  MoveL 521 to (0, -31.79, 55.65) mm, rotated rx 170.45 ry 0 rz 180 deg; joints [-13.216, -55.69, 111.554, 164.16, 56.887, -90.738]
  MoveL 522 to (-200, -31.79, 55.65) mm, rotated rx 170.45 ry 0 rz 180 deg; joints [-15.372, -64.732, 127.633, 162.838, 63.944, -91.824]
  MoveL 523 to (-200, -32.38, 55.53) mm, rotated rx 167.27 ry 0 rz 180 deg; joints [-15.299, -65.985, 127.45, 162.704, 62.564, -94.567]
  MoveL 524 to (0, -32.38, 55.53) mm, rotated rx 167.27 ry 0 rz 180 deg; joints [-13.153, -56.711, 111.391, 164.018, 55.738, -93.573]
  MoveL 525 to (0, -32.96, 55.39) mm, rotated rx 164.09 ry 0 rz 180 deg; joints [-13.044, -57.718, 111.217, 163.922, 54.585, -96.433]
  MoveL 526 to (-200, -32.96, 55.39) mm, rotated rx 164.09 ry 0 rz 180 deg; joints [-15.175, -67.219, 127.255, 162.616, 61.181, -97.333]
  MoveL 527 to (-200, -33.53, 55.21) mm, rotated rx 160.9 ry 0 rz 180 deg; joints [-14.999, -68.432, 127.047, 162.576, 59.799, -100.128]
  MoveL 528 to (0, -33.53, 55.21) mm, rotated rx 160.9 ry 0 rz 180 deg; joints [-12.891, -58.708, 111.032, 163.872, 53.431, -99.324]
  MoveL 529 to (0, -34.09, 54.99) mm, rotated rx 157.72 ry 0 rz 180 deg; joints [-12.693, -59.678, 110.838, 163.872, 52.279, -102.249]
  MoveL 530 to (-200, -34.09, 54.99) mm, rotated rx 157.72 ry 0 rz 180 deg; joints [-14.771, -69.618, 126.828, 162.586, 58.422, -102.955]
  MoveL 531 to (-200, -34.64, 54.75) mm, rotated rx 154.53 ry 0 rz 180 deg; joints [-14.492, -70.775, 126.599, 162.65, 57.053, -105.822]
  MoveL 532 to (0, -34.64, 54.75) mm, rotated rx 154.53 ry 0 rz 180 deg; joints [-12.451, -60.626, 110.636, 163.924, 51.131, -105.214]
  MoveL 533 to (0, -35.18, 54.48) mm, rotated rx 151.35 ry 0 rz 180 deg; joints [-12.165, -61.547, 110.426, 164.031, 49.993, -108.224]
  MoveL 534 to (-200, -35.18, 54.48) mm, rotated rx 151.35 ry 0 rz 180 deg; joints [-14.163, -71.9, 126.361, 162.77, 55.696, -108.734]
  MoveL 535 to (-200, -35.7, 54.18) mm, rotated rx 148.17 ry 0 rz 180 deg; joints [-13.784, -72.989, 126.115, 162.95, 54.354, -111.698]
  MoveL 536 to (0, -35.7, 54.18) mm, rotated rx 148.17 ry 0 rz 180 deg; joints [-11.836, -62.442, 110.21, 164.197, 48.865, -111.284]
  MoveL 537 to (0, -36.2, 53.84) mm, rotated rx 144.99 ry 0 rz 180 deg; joints [-11.464, -63.305, 109.989, 164.425, 47.752, -114.399]
  MoveL 538 to (-200, -36.2, 53.84) mm, rotated rx 144.99 ry 0 rz 180 deg; joints [-13.356, -74.041, 125.863, 163.195, 53.031, -114.72]
  MoveL 539 to (-200, -36.68, 53.49) mm, rotated rx 141.8 ry 0 rz 180 deg; joints [-12.879, -75.052, 125.607, 163.507, 51.731, -117.806]
  MoveL 540 to (0, -36.68, 53.49) mm, rotated rx 141.8 ry 0 rz 180 deg; joints [-11.052, -64.137, 109.764, 164.717, 46.658, -117.575]
  MoveL 541 to (0, -37.14, 53.1) mm, rotated rx 138.62 ry 0 rz 180 deg; joints [-10.598, -64.933, 109.536, 165.079, 45.585, -120.816]
  MoveL 542 to (-200, -37.14, 53.1) mm, rotated rx 138.62 ry 0 rz 180 deg; joints [-12.355, -76.019, 125.348, 163.891, 50.459, -120.962]
  MoveL 543 to (-200, -37.58, 52.7) mm, rotated rx 135.44 ry 0 rz 180 deg; joints [-11.785, -76.941, 125.087, 164.352, 49.218, -124.195]
  MoveL 544 to (0, -37.58, 52.7) mm, rotated rx 135.44 ry 0 rz 180 deg; joints [-10.105, -65.693, 109.307, 165.513, 44.539, -124.128]
  MoveL 545 to (0, -37.99, 52.26) mm, rotated rx 132.25 ry 0 rz 180 deg; joints [-9.574, -66.415, 109.079, 166.023, 43.523, -127.516]
  MoveL 546 to (-200, -37.99, 52.26) mm, rotated rx 132.25 ry 0 rz 180 deg; joints [-11.17, -77.816, 124.826, 164.893, 48.014, -127.51]
  MoveL 547 to (-200, -38.38, 51.81) mm, rotated rx 129.07 ry 0 rz 180 deg; joints [-10.512, -78.64, 124.568, 165.519, 46.851, -130.914]
  MoveL 548 to (0, -38.38, 51.81) mm, rotated rx 129.07 ry 0 rz 180 deg; joints [-9.006, -67.096, 108.852, 166.613, 42.541, -130.984]
  MoveL 549 to (0, -38.75, 51.33) mm, rotated rx 125.89 ry 0 rz 180 deg; joints [-8.403, -67.735, 108.628, 167.284, 41.598, -134.535]
  MoveL 550 to (-200, -38.75, 51.33) mm, rotated rx 125.89 ry 0 rz 180 deg; joints [-9.811, -79.413, 124.313, 166.234, 45.735, -134.409]
  MoveL 551 to (-200, -39.09, 50.84) mm, rotated rx 122.7 ry 0 rz 180 deg; joints [-9.071, -80.133, 124.064, 167.04, 44.67, -138.001]
  MoveL 552 to (0, -39.09, 50.84) mm, rotated rx 122.7 ry 0 rz 180 deg; joints [-7.766, -68.33, 108.408, 168.04, 40.698, -138.172]
  MoveL 553 to (0, -39.4, 50.32) mm, rotated rx 119.52 ry 0 rz 180 deg; joints [-7.098, -68.881, 108.194, 168.881, 39.847, -141.898]
  MoveL 554 to (-200, -39.4, 50.32) mm, rotated rx 119.52 ry 0 rz 180 deg; joints [-8.293, -80.797, 123.822, 167.941, 43.662, -141.693]
  MoveL 555 to (-200, -39.68, 49.79) mm, rotated rx 116.34 ry 0 rz 180 deg; joints [-7.48, -81.406, 123.588, 168.937, 42.718, -145.487]
  MoveL 556 to (0, -39.68, 49.79) mm, rotated rx 116.34 ry 0 rz 180 deg; joints [-6.399, -69.385, 107.988, 169.809, 39.048, -145.714]
  MoveL 557 to (0, -39.93, 49.25) mm, rotated rx 113.16 ry 0 rz 180 deg; joints [-5.673, -69.842, 107.79, 170.823, 38.306, -149.62]
  MoveL 558 to (-200, -39.93, 49.25) mm, rotated rx 113.16 ry 0 rz 180 deg; joints [-6.633, -81.956, 123.364, 170.028, 41.841, -149.382]
  MoveL 559 to (-200, -40.15, 48.69) mm, rotated rx 109.97 ry 0 rz 180 deg; joints [-5.756, -82.448, 123.153, 171.213, 41.039, -153.378]
  MoveL 560 to (0, -40.15, 48.69) mm, rotated rx 109.97 ry 0 rz 180 deg; joints [-4.922, -70.251, 107.602, 171.922, 37.627, -153.614]
  MoveL 561 to (0, -40.34, 48.12) mm, rotated rx 106.79 ry 0 rz 180 deg; joints [-4.147, -70.61, 107.424, 173.101, 37.014, -157.692]
  MoveL 562 to (-200, -40.34, 48.12) mm, rotated rx 106.79 ry 0 rz 180 deg; joints [-4.852, -82.881, 122.954, 172.489, 40.317, -157.47]
  MoveL 563 to (-200, -40.5, 47.54) mm, rotated rx 103.61 ry 0 rz 180 deg; joints [-3.922, -83.252, 122.77, 173.85, 39.68, -161.653]
  MoveL 564 to (0, -40.5, 47.54) mm, rotated rx 103.61 ry 0 rz 180 deg; joints [-3.352, -70.919, 107.259, 174.355, 36.473, -161.85]
  MoveL 565 to (0, -40.62, 46.95) mm, rotated rx 100.42 ry 0 rz 180 deg; joints [-2.539, -71.178, 107.107, 175.679, 36.006, -166.079]
  MoveL 566 to (-200, -40.62, 46.95) mm, rotated rx 100.42 ry 0 rz 180 deg; joints [-2.971, -83.563, 122.601, 175.289, 39.133, -165.919]
  MoveL 567 to (-200, -40.71, 46.36) mm, rotated rx 97.24 ry 0 rz 180 deg; joints [-2.002, -83.812, 122.449, 176.795, 38.681, -170.258]
  MoveL 568 to (0, -40.71, 46.36) mm, rotated rx 97.24 ry 0 rz 180 deg; joints [-1.711, -71.386, 106.969, 177.062, 35.619, -170.372]
  MoveL 569 to (0, -40.77, 45.76) mm, rotated rx 94.06 ry 0 rz 180 deg; joints [-0.87, -71.542, 106.846, 178.494, 35.313, -174.715]
  MoveL 570 to (-200, -40.77, 45.76) mm, rotated rx 94.06 ry 0 rz 180 deg; joints [-1.019, -83.999, 122.314, 178.357, 38.327, -174.655]
  MoveL 571 to (-200, -40.8, 45.16) mm, rotated rx 90.87 ry 0 rz 180 deg; joints [-0.024, -84.123, 122.198, 179.961, 38.074, -179.096]
  MoveL 572 to (0, -40.8, 45.16) mm, rotated rx 90.87 ry 0 rz 180 deg; joints [-0.021, -71.646, 106.738, 179.964, 35.092, -179.097]
  MoveL 573 to (0, -40.8, 44.56) mm, rotated rx 90 ry 0 rz 180 deg; joints [0.232, -71.666, 106.711, -179.597, 35.046, 179.67]
  MoveL 574 to (-200, -40.8, 44.56) mm, rotated rx 90 ry 0 rz 180 deg; joints [0.271, -84.147, 122.169, -179.56, 38.023, 179.653]
  MoveL 575 to (-200, -40.8, 43.97) mm, rotated rx 90 ry 0 rz 180 deg; joints [0.301, -84.146, 122.169, -179.512, 38.023, 179.616]
  MoveL 576 to (0, -40.8, 43.97) mm, rotated rx 90 ry 0 rz 180 deg; joints [0.257, -71.666, 106.711, -179.553, 35.046, 179.634]
  MoveL 577 to (0, -40.8, 43.37) mm, rotated rx 90 ry 0 rz 180 deg; joints [0.282, -71.665, 106.711, -179.509, 35.046, 179.598]
  MoveL 578 to (-200, -40.8, 43.37) mm, rotated rx 90 ry 0 rz 180 deg; joints [0.33, -84.146, 122.169, -179.464, 38.024, 179.578]
  MoveL 579 to (-200, -40.8, 42.77) mm, rotated rx 90 ry 0 rz 180 deg; joints [0.359, -84.146, 122.168, -179.417, 38.024, 179.541]
  MoveL 580 to (0, -40.8, 42.77) mm, rotated rx 90 ry 0 rz 180 deg; joints [0.307, -71.665, 106.71, -179.466, 35.046, 179.562]
  MoveL 581 to (0, -40.8, 42.16) mm, rotated rx 90 ry 0 rz 180 deg; joints [0.332, -71.665, 106.71, -179.422, 35.046, 179.527]
  MoveL 582 to (-200, -40.8, 42.16) mm, rotated rx 90 ry 0 rz 180 deg; joints [0.389, -84.146, 122.168, -179.369, 38.024, 179.503]
  MoveL 583 to (-200, -40.8, 41.56) mm, rotated rx 90 ry 0 rz 180 deg; joints [0.418, -84.145, 122.168, -179.322, 38.024, 179.466]
  MoveL 584 to (0, -40.8, 41.56) mm, rotated rx 90 ry 0 rz 180 deg; joints [0.357, -71.665, 106.71, -179.378, 35.047, 179.491]
  MoveL 585 to (0, -40.8, 40.97) mm, rotated rx 90 ry 0 rz 180 deg; joints [0.382, -71.665, 106.709, -179.335, 35.047, 179.455]
  MoveL 586 to (-200, -40.8, 40.97) mm, rotated rx 90 ry 0 rz 180 deg; joints [0.447, -84.145, 122.167, -179.274, 38.025, 179.428]
  MoveL 587 to (-200, -40.8, 40.37) mm, rotated rx 90 ry 0 rz 180 deg; joints [0.477, -84.145, 122.167, -179.226, 38.025, 179.391]
  MoveL 588 to (0, -40.8, 40.37) mm, rotated rx 90 ry 0 rz 180 deg; joints [0.407, -71.664, 106.709, -179.291, 35.047, 179.42]
  MoveL 589 to (0, -40.8, 39.77) mm, rotated rx 90 ry 0 rz 180 deg; joints [0.432, -71.664, 106.709, -179.247, 35.047, 179.384]
  MoveL 590 to (-200, -40.8, 39.77) mm, rotated rx 90 ry 0 rz 180 deg; joints [0.506, -84.144, 122.167, -179.179, 38.025, 179.353]
  MoveL 591 to (-200, -40.8, 39.16) mm, rotated rx 90 ry 0 rz 180 deg; joints [0.535, -84.144, 122.166, -179.131, 38.025, 179.316]
  MoveL 592 to (0, -40.8, 39.16) mm, rotated rx 90 ry 0 rz 180 deg; joints [0.457, -71.664, 106.708, -179.204, 35.047, 179.348]
  MoveL 593 to (0, -40.8, 38.56) mm, rotated rx 90 ry 0 rz 180 deg; joints [0.482, -71.663, 106.708, -179.16, 35.047, 179.312]
  MoveL 594 to (-200, -40.8, 38.56) mm, rotated rx 90 ry 0 rz 180 deg; joints [0.565, -84.144, 122.166, -179.084, 38.026, 179.278]
  MoveL 595 to (-200, -40.8, 37.97) mm, rotated rx 90 ry 0 rz 180 deg; joints [0.594, -84.143, 122.165, -179.036, 38.026, 179.241]
  MoveL 596 to (0, -40.8, 37.97) mm, rotated rx 90 ry 0 rz 180 deg; joints [0.507, -71.663, 106.708, -179.117, 35.048, 179.277]
  MoveL 597 to (0, -40.8, 37.37) mm, rotated rx 90 ry 0 rz 180 deg; joints [0.532, -71.663, 106.707, -179.073, 35.048, 179.241]
  MoveL 598 to (-200, -40.8, 37.37) mm, rotated rx 90 ry 0 rz 180 deg; joints [0.623, -84.143, 122.165, -178.988, 38.026, 179.203]
  MoveL 599 to (-200, -40.8, 36.77) mm, rotated rx 90 ry 0 rz 180 deg; joints [0.653, -84.143, 122.165, -178.941, 38.027, 179.166]
  MoveL 600 to (0, -40.8, 36.77) mm, rotated rx 90 ry 0 rz 180 deg; joints [0.557, -71.662, 106.707, -179.029, 35.048, 179.205]
  MoveL 601 to (0, -40.8, 36.16) mm, rotated rx 90 ry 0 rz 180 deg; joints [0.582, -71.662, 106.706, -178.986, 35.048, 179.17]
  MoveL 602 to (-200, -40.8, 36.16) mm, rotated rx 90 ry 0 rz 180 deg; joints [0.682, -84.142, 122.164, -178.893, 38.027, 179.128]
  MoveL 603 to (-200, -40.8, 35.56) mm, rotated rx 90 ry 0 rz 180 deg; joints [0.711, -84.142, 122.163, -178.845, 38.028, 179.091]
  MoveL 604 to (0, -40.8, 35.56) mm, rotated rx 90 ry 0 rz 180 deg; joints [0.608, -71.662, 106.706, -178.942, 35.048, 179.134]
  MoveL 605 to (0, -40.8, 34.97) mm, rotated rx 90 ry 0 rz 180 deg; joints [0.633, -71.661, 106.705, -178.898, 35.049, 179.098]
  MoveL 606 to (-200, -40.8, 34.97) mm, rotated rx 90 ry 0 rz 180 deg; joints [0.741, -84.141, 122.163, -178.798, 38.028, 179.053]
  MoveL 607 to (-200, -40.8, 34.37) mm, rotated rx 90 ry 0 rz 180 deg; joints [0.77, -84.141, 122.162, -178.75, 38.028, 179.016]
  MoveL 608 to (0, -40.8, 34.37) mm, rotated rx 90 ry 0 rz 180 deg; joints [0.658, -71.661, 106.704, -178.855, 35.049, 179.062]
  MoveL 609 to (0, -40.8, 33.77) mm, rotated rx 90 ry 0 rz 180 deg; joints [0.683, -71.66, 106.704, -178.811, 35.049, 179.027]
  MoveL 610 to (-200, -40.8, 33.77) mm, rotated rx 90 ry 0 rz 180 deg; joints [0.799, -84.14, 122.162, -178.703, 38.029, 178.978]
  MoveL 611 to (-200, -40.8, 33.16) mm, rotated rx 90 ry 0 rz 180 deg; joints [0.829, -84.14, 122.161, -178.655, 38.029, 178.941]
  MoveL 612 to (0, -40.8, 33.16) mm, rotated rx 90 ry 0 rz 180 deg; joints [0.708, -71.66, 106.703, -178.768, 35.05, 178.991]
  MoveL 613 to (0, -40.8, 32.56) mm, rotated rx 90 ry 0 rz 180 deg; joints [0.733, -71.66, 106.703, -178.724, 35.05, 178.955]
  MoveL 614 to (-200, -40.8, 32.56) mm, rotated rx 90 ry 0 rz 180 deg; joints [0.858, -84.139, 122.161, -178.607, 38.03, 178.903]
  MoveL 615 to (-200, -40.8, 31.96) mm, rotated rx 90 ry 0 rz 180 deg; joints [0.887, -84.138, 122.16, -178.56, 38.03, 178.866]
  MoveL 616 to (0, -40.8, 31.96) mm, rotated rx 90 ry 0 rz 180 deg; joints [0.758, -71.659, 106.702, -178.68, 35.05, 178.92]
  MoveL 617 to (0, -40.8, 31.36) mm, rotated rx 90 ry 0 rz 180 deg; joints [0.783, -71.659, 106.701, -178.637, 35.05, 178.884]
  MoveL 618 to (-200, -40.8, 31.36) mm, rotated rx 90 ry 0 rz 180 deg; joints [0.916, -84.138, 122.159, -178.512, 38.031, 178.828]
  MoveL 619 to (-200, -40.8, 30.77) mm, rotated rx 90 ry 0 rz 180 deg; joints [0.946, -84.137, 122.158, -178.465, 38.031, 178.791]
  MoveL 620 to (0, -40.8, 30.77) mm, rotated rx 90 ry 0 rz 180 deg; joints [0.808, -71.658, 106.701, -178.593, 35.051, 178.848]
  MoveL 621 to (0, -40.8, 30.16) mm, rotated rx 90 ry 0 rz 180 deg; joints [0.833, -71.657, 106.7, -178.549, 35.051, 178.812]
  MoveL 622 to (-200, -40.8, 30.16) mm, rotated rx 90 ry 0 rz 180 deg; joints [0.975, -84.136, 122.158, -178.417, 38.032, 178.753]
  MoveL 623 to (-200, -40.8, 29.57) mm, rotated rx 90 ry 0 rz 180 deg; joints [1.004, -84.136, 122.157, -178.37, 38.032, 178.716]
  MoveL 624 to (0, -40.8, 29.57) mm, rotated rx 90 ry 0 rz 180 deg; joints [0.858, -71.657, 106.699, -178.506, 35.051, 178.777]
  MoveL 625 to (0, -40.8, 28.96) mm, rotated rx 90 ry 0 rz 180 deg; joints [0.883, -71.656, 106.698, -178.462, 35.052, 178.741]
  MoveL 626 to (-200, -40.8, 28.96) mm, rotated rx 90 ry 0 rz 180 deg; joints [1.034, -84.135, 122.156, -178.322, 38.033, 178.678]
  MoveL 627 to (-200, -40.8, 28.36) mm, rotated rx 90 ry 0 rz 180 deg; joints [1.063, -84.134, 122.155, -178.274, 38.034, 178.641]
  MoveL 628 to (0, -40.8, 28.36) mm, rotated rx 90 ry 0 rz 180 deg; joints [0.908, -71.656, 106.698, -178.419, 35.052, 178.705]
  MoveL 629 to (0, -40.8, 27.77) mm, rotated rx 90 ry 0 rz 180 deg; joints [0.933, -71.655, 106.697, -178.375, 35.052, 178.67]
  MoveL 630 to (-200, -40.8, 27.77) mm, rotated rx 90 ry 0 rz 180 deg; joints [1.092, -84.134, 122.155, -178.227, 38.034, 178.603]
  MoveL 631 to (-200, -40.8, 27.16) mm, rotated rx 90 ry 0 rz 180 deg; joints [1.122, -84.133, 122.154, -178.179, 38.035, 178.566]
  MoveL 632 to (0, -40.8, 27.16) mm, rotated rx 90 ry 0 rz 180 deg; joints [0.958, -71.655, 106.696, -178.331, 35.053, 178.634]
  MoveL 633 to (0, -40.8, 26.57) mm, rotated rx 90 ry 0 rz 180 deg; joints [0.983, -71.654, 106.695, -178.288, 35.053, 178.598]
  MoveL 634 to (-200, -40.8, 26.57) mm, rotated rx 90 ry 0 rz 180 deg; joints [1.151, -84.132, 122.153, -178.132, 38.036, 178.528]
  MoveL 635 to (-200, -40.8, 25.96) mm, rotated rx 90 ry 0 rz 180 deg; joints [1.18, -84.131, 122.152, -178.084, 38.036, 178.491]
  MoveL 636 to (0, -40.8, 25.96) mm, rotated rx 90 ry 0 rz 180 deg; joints [1.008, -71.653, 106.694, -178.244, 35.054, 178.562]
  MoveL 637 to (0, -40.8, 25.36) mm, rotated rx 90 ry 0 rz 180 deg; joints [1.033, -71.653, 106.693, -178.201, 35.054, 178.527]
  MoveL 638 to (-200, -40.8, 25.36) mm, rotated rx 90 ry 0 rz 180 deg; joints [1.21, -84.131, 122.151, -178.036, 38.037, 178.453]
  MoveL 639 to (-200, -40.8, 24.77) mm, rotated rx 90 ry 0 rz 180 deg; joints [1.239, -84.13, 122.15, -177.989, 38.038, 178.416]
  MoveL 640 to (0, -40.8, 24.77) mm, rotated rx 90 ry 0 rz 180 deg; joints [1.058, -71.652, 106.692, -178.157, 35.054, 178.491]
  MoveL 641 to (0, -40.8, 24.16) mm, rotated rx 90 ry 0 rz 180 deg; joints [1.084, -71.651, 106.692, -178.113, 35.055, 178.455]
  MoveL 642 to (-200, -40.8, 24.16) mm, rotated rx 90 ry 0 rz 180 deg; joints [1.268, -84.129, 122.149, -177.941, 38.038, 178.378]
  MoveL 643 to (-200, -40.8, 23.57) mm, rotated rx 90 ry 0 rz 180 deg; joints [1.298, -84.128, 122.148, -177.894, 38.039, 178.341]
  MoveL 644 to (0, -40.8, 23.57) mm, rotated rx 90 ry 0 rz 180 deg; joints [1.109, -71.651, 106.691, -178.07, 35.055, 178.42]
  MoveL 645 to (0, -40.8, 22.96) mm, rotated rx 90 ry 0 rz 180 deg; joints [1.134, -71.65, 106.69, -178.026, 35.056, 178.384]
  MoveL 646 to (-200, -40.8, 22.96) mm, rotated rx 90 ry 0 rz 180 deg; joints [1.327, -84.127, 122.147, -177.846, 38.04, 178.303]
  MoveL 647 to (-200, -40.8, 22.36) mm, rotated rx 90 ry 0 rz 180 deg; joints [1.356, -84.126, 122.146, -177.799, 38.041, 178.266]
  MoveL 648 to (0, -40.8, 22.36) mm, rotated rx 90 ry 0 rz 180 deg; joints [1.159, -71.649, 106.689, -177.982, 35.056, 178.348]
  MoveL 649 to (0, -40.8, 21.77) mm, rotated rx 90 ry 0 rz 180 deg; joints [1.184, -71.648, 106.688, -177.939, 35.057, 178.313]
  MoveL 650 to (-200, -40.8, 21.77) mm, rotated rx 90 ry 0 rz 180 deg; joints [1.386, -84.125, 122.145, -177.751, 38.041, 178.228]
  MoveL 651 to (-200, -40.8, 21.16) mm, rotated rx 90 ry 0 rz 180 deg; joints [1.415, -84.124, 122.144, -177.704, 38.042, 178.191]
  MoveL 652 to (0, -40.8, 21.16) mm, rotated rx 90 ry 0 rz 180 deg; joints [1.209, -71.648, 106.687, -177.895, 35.057, 178.277]
  MoveL 653 to (0, -40.8, 20.57) mm, rotated rx 90 ry 0 rz 180 deg; joints [1.234, -71.647, 106.685, -177.852, 35.058, 178.241]
  MoveL 654 to (-200, -40.8, 20.57) mm, rotated rx 90 ry 0 rz 180 deg; joints [1.444, -84.123, 122.143, -177.656, 38.043, 178.154]
  MoveL 655 to (-200, -40.8, 19.96) mm, rotated rx 90 ry 0 rz 180 deg; joints [1.474, -84.122, 122.142, -177.608, 38.044, 178.116]
  MoveL 656 to (0, -40.8, 19.96) mm, rotated rx 90 ry 0 rz 180 deg; joints [1.259, -71.646, 106.684, -177.808, 35.058, 178.205]
  MoveL 657 to (0, -40.8, 19.36) mm, rotated rx 90 ry 0 rz 180 deg; joints [1.284, -71.645, 106.683, -177.765, 35.059, 178.17]
  MoveL 658 to (-200, -40.8, 19.36) mm, rotated rx 90 ry 0 rz 180 deg; joints [1.503, -84.121, 122.141, -177.561, 38.045, 178.079]
  MoveL 659 to (-200, -40.8, 18.77) mm, rotated rx 90 ry 0 rz 180 deg; joints [1.532, -84.12, 122.14, -177.513, 38.046, 178.041]
  MoveL 660 to (0, -40.8, 18.77) mm, rotated rx 90 ry 0 rz 180 deg; joints [1.309, -71.644, 106.682, -177.721, 35.059, 178.134]
  MoveL 661 to (0, -40.8, 18.16) mm, rotated rx 90 ry 0 rz 180 deg; joints [1.334, -71.644, 106.681, -177.677, 35.06, 178.098]
  MoveL 662 to (-200, -40.8, 18.16) mm, rotated rx 90 ry 0 rz 180 deg; joints [1.562, -84.119, 122.139, -177.466, 38.046, 178.004]
  MoveL 663 to (-200, -40.8, 17.57) mm, rotated rx 90 ry 0 rz 180 deg; joints [1.591, -84.118, 122.137, -177.418, 38.047, 177.966]
  MoveL 664 to (0, -40.8, 17.57) mm, rotated rx 90 ry 0 rz 180 deg; joints [1.359, -71.643, 106.68, -177.634, 35.06, 178.063]
  MoveL 665 to (0, -40.8, 16.96) mm, rotated rx 90 ry 0 rz 180 deg; joints [1.384, -71.642, 106.679, -177.59, 35.061, 178.027]
  MoveL 666 to (-200, -40.8, 16.96) mm, rotated rx 90 ry 0 rz 180 deg; joints [1.62, -84.117, 122.136, -177.371, 38.048, 177.929]
  MoveL 667 to (-200, -40.8, 16.36) mm, rotated rx 90 ry 0 rz 180 deg; joints [1.649, -84.116, 122.135, -177.323, 38.049, 177.891]
  MoveL 668 to (0, -40.8, 16.36) mm, rotated rx 90 ry 0 rz 180 deg; joints [1.409, -71.641, 106.677, -177.547, 35.061, 177.991]
  MoveL 669 to (0, -40.8, 15.77) mm, rotated rx 90 ry 0 rz 180 deg; joints [1.434, -71.64, 106.676, -177.503, 35.062, 177.956]
  MoveL 670 to (-200, -40.8, 15.77) mm, rotated rx 90 ry 0 rz 180 deg; joints [1.679, -84.115, 122.134, -177.276, 38.05, 177.854]
  MoveL 671 to (-200, -40.8, 15.16) mm, rotated rx 90 ry 0 rz 180 deg; joints [1.708, -84.114, 122.133, -177.228, 38.051, 177.817]
  MoveL 672 to (0, -40.8, 15.16) mm, rotated rx 90 ry 0 rz 180 deg; joints [1.459, -71.639, 106.675, -177.459, 35.062, 177.92]
  MoveL 673 to (0, -40.79, 14.56) mm, rotated rx 87.69 ry 0 rz 180 deg; joints [2.087, -71.652, 106.583, -176.358, 34.985, 174.705]
  MoveL 674 to (-200, -40.79, 14.56) mm, rotated rx 87.69 ry 0 rz 180 deg; joints [2.443, -84.128, 122.036, -176.028, 37.975, 174.557]
  MoveL 675 to (-200, -40.75, 13.97) mm, rotated rx 84.51 ry 0 rz 180 deg; joints [3.447, -84.094, 121.92, -174.391, 37.959, 170.079]
  MoveL 676 to (0, -40.75, 13.97) mm, rotated rx 84.51 ry 0 rz 180 deg; joints [2.945, -71.625, 106.47, -174.855, 34.954, 170.286]
  MoveL 677 to (0, -40.68, 13.37) mm, rotated rx 81.32 ry 0 rz 180 deg; joints [3.803, -71.546, 106.374, -173.362, 35.009, 165.879]
  MoveL 678 to (-200, -40.68, 13.37) mm, rotated rx 81.32 ry 0 rz 180 deg; joints [4.449, -83.998, 121.824, -172.769, 38.047, 165.618]
  MoveL 679 to (-200, -40.57, 12.78) mm, rotated rx 78.14 ry 0 rz 180 deg; joints [5.447, -83.841, 121.747, -171.177, 38.237, 161.19]
  MoveL 680 to (0, -40.57, 12.78) mm, rotated rx 78.14 ry 0 rz 180 deg; joints [4.657, -71.416, 106.295, -171.893, 35.15, 161.498]
  MoveL 681 to (0, -40.43, 12.2) mm, rotated rx 74.96 ry 0 rz 180 deg; joints [5.505, -71.235, 106.233, -170.462, 35.374, 157.157]
  MoveL 682 to (-200, -40.43, 12.2) mm, rotated rx 74.96 ry 0 rz 180 deg; joints [6.437, -83.622, 121.69, -169.631, 38.527, 156.812]
  MoveL 683 to (-200, -40.26, 11.62) mm, rotated rx 71.78 ry 0 rz 180 deg; joints [7.415, -83.344, 121.653, -168.144, 38.911, 152.498]
  MoveL 684 to (0, -40.26, 11.62) mm, rotated rx 71.78 ry 0 rz 180 deg; joints [6.343, -71.004, 106.189, -169.08, 35.679, 152.868]
  MoveL 685 to (0, -40.05, 11.06) mm, rotated rx 68.59 ry 0 rz 180 deg; joints [7.17, -70.724, 106.161, -167.759, 36.062, 148.644]
  MoveL 686 to (-200, -40.05, 11.06) mm, rotated rx 68.59 ry 0 rz 180 deg; joints [8.377, -83.007, 121.635, -166.727, 39.387, 148.26]
  MoveL 687 to (-200, -39.82, 10.51) mm, rotated rx 65.41 ry 0 rz 180 deg; joints [9.322, -82.611, 121.637, -165.389, 39.95, 144.107]
  MoveL 688 to (0, -39.82, 10.51) mm, rotated rx 65.41 ry 0 rz 180 deg; joints [7.982, -70.395, 106.15, -166.506, 36.518, 144.492]
  MoveL 689 to (0, -39.56, 9.97) mm, rotated rx 62.22 ry 0 rz 180 deg; joints [8.776, -70.019, 106.155, -165.33, 37.045, 140.423]
  MoveL 690 to (-200, -39.56, 9.97) mm, rotated rx 62.22 ry 0 rz 180 deg; joints [10.244, -82.159, 121.657, -164.139, 40.593, 140.05]
  MoveL 691 to (-200, -39.26, 9.44) mm, rotated rx 59.04 ry 0 rz 180 deg; joints [11.141, -81.651, 121.694, -162.98, 41.312, 136.093]
  MoveL 692 to (0, -39.26, 9.44) mm, rotated rx 59.04 ry 0 rz 180 deg; joints [9.55, -69.596, 106.175, -164.236, 37.636, 136.441]
  MoveL 693 to (0, -38.94, 8.94) mm, rotated rx 55.86 ry 0 rz 180 deg; joints [10.301, -69.128, 106.211, -163.226, 38.289, 132.549]
  MoveL 694 to (-200, -38.94, 8.94) mm, rotated rx 55.86 ry 0 rz 180 deg; joints [12.011, -81.089, 121.748, -161.916, 42.099, 132.239]
  MoveL 695 to (-200, -38.59, 8.45) mm, rotated rx 52.68 ry 0 rz 180 deg; joints [12.851, -80.474, 121.819, -160.948, 42.951, 128.49]
  MoveL 696 to (0, -38.59, 8.45) mm, rotated rx 52.68 ry 0 rz 180 deg; joints [11.028, -68.615, 106.262, -162.304, 38.997, 128.749]
  MoveL 697 to (0, -38.21, 7.99) mm, rotated rx 49.49 ry 0 rz 180 deg; joints [11.727, -68.06, 106.326, -161.469, 39.757, 125.043]
  MoveL 698 to (-200, -38.21, 7.99) mm, rotated rx 49.49 ry 0 rz 180 deg; joints [13.659, -79.807, 121.905, -160.075, 43.861, 124.846]
  MoveL 699 to (-200, -37.81, 7.54) mm, rotated rx 46.31 ry 0 rz 180 deg; joints [14.431, -79.092, 122.004, -159.296, 44.823, 121.303]
  MoveL 700 to (0, -37.81, 7.54) mm, rotated rx 46.31 ry 0 rz 180 deg; joints [12.398, -67.464, 106.403, -160.722, 40.564, 121.43]
  MoveL 701 to (0, -37.38, 7.12) mm, rotated rx 43.13 ry 0 rz 180 deg; joints [13.038, -66.828, 106.491, -160.059, 41.413, 117.906]
  MoveL 702 to (-200, -37.38, 7.12) mm, rotated rx 43.13 ry 0 rz 180 deg; joints [15.167, -78.328, 122.117, -158.608, 45.833, 117.86]
  MoveL 703 to (-200, -36.93, 6.72) mm, rotated rx 39.94 ry 0 rz 180 deg; joints [15.865, -77.519, 122.241, -158.007, 46.885, 114.512]
  MoveL 704 to (0, -36.93, 6.72) mm, rotated rx 39.94 ry 0 rz 180 deg; joints [13.646, -66.153, 106.591, -159.48, 42.3, 114.47]
  MoveL 705 to (0, -36.46, 6.35) mm, rotated rx 36.76 ry 0 rz 180 deg; joints [14.219, -65.442, 106.7, -158.98, 43.221, 111.118]
  MoveL 706 to (-200, -36.46, 6.35) mm, rotated rx 36.76 ry 0 rz 180 deg; joints [16.522, -76.665, 122.375, -157.49, 47.975, 111.255]
  MoveL 707 to (-200, -35.97, 6) mm, rotated rx 33.58 ry 0 rz 180 deg; joints [17.139, -75.77, 122.519, -157.053, 49.098, 108.083]
  MoveL 708 to (0, -35.97, 6) mm, rotated rx 33.58 ry 0 rz 180 deg; joints [14.758, -64.697, 106.818, -158.557, 44.172, 107.844]
  MoveL 709 to (0, -35.46, 5.68) mm, rotated rx 30.39 ry 0 rz 180 deg; joints [15.259, -63.918, 106.944, -158.208, 45.149, 104.647]
  MoveL 710 to (-200, -35.46, 5.68) mm, rotated rx 30.39 ry 0 rz 180 deg; joints [17.712, -74.835, 122.67, -156.691, 50.25, 104.99]
  MoveL 711 to (-200, -34.94, 5.39) mm, rotated rx 27.21 ry 0 rz 180 deg; joints [18.241, -73.862, 122.828, -156.399, 51.427, 101.972]
  MoveL 712 to (0, -34.94, 5.39) mm, rotated rx 27.21 ry 0 rz 180 deg; joints [15.723, -63.109, 107.077, -157.927, 46.149, 101.519]
  MoveL 713 to (0, -34.4, 5.14) mm, rotated rx 24.03 ry 0 rz 180 deg; joints [16.149, -62.27, 107.216, -157.712, 47.168, 98.457]
  MoveL 714 to (-200, -34.4, 5.14) mm, rotated rx 24.03 ry 0 rz 180 deg; joints [18.725, -72.854, 122.992, -156.174, 52.626, 99.022]
  MoveL 715 to (-200, -33.84, 4.91) mm, rotated rx 20.84 ry 0 rz 180 deg; joints [19.164, -71.813, 123.16, -156.01, 53.843, 96.134]
  MoveL 716 to (0, -33.84, 4.91) mm, rotated rx 20.84 ry 0 rz 180 deg; joints [16.534, -61.405, 107.359, -157.559, 48.203, 95.454]
  MoveL 717 to (0, -33.28, 4.71) mm, rotated rx 17.66 ry 0 rz 180 deg; joints [16.88, -60.515, 107.506, -157.463, 49.252, 92.507]
  MoveL 718 to (-200, -33.28, 4.71) mm, rotated rx 17.66 ry 0 rz 180 deg; joints [19.556, -70.742, 123.33, -155.905, 55.076, 93.301]
  MoveL 719 to (-200, -32.7, 4.54) mm, rotated rx 14.48 ry 0 rz 180 deg; joints [19.901, -69.642, 123.503, -155.854, 56.322, 90.519]
  MoveL 720 to (0, -32.7, 4.54) mm, rotated rx 14.48 ry 0 rz 180 deg; joints [17.184, -59.603, 107.655, -157.423, 50.312, 89.608]
  MoveL 721 to (0, -32.12, 4.41) mm, rotated rx 11.3 ry 0 rz 180 deg; joints [17.447, -58.67, 107.807, -157.434, 51.38, 86.755]
  MoveL 722 to (-200, -32.12, 4.41) mm, rotated rx 11.3 ry 0 rz 180 deg; joints [20.199, -68.517, 123.676, -155.855, 57.577, 87.781]
  MoveL 723 to (-200, -31.52, 4.31) mm, rotated rx 8.11 ry 0 rz 180 deg; joints [20.449, -67.37, 123.849, -155.903, 58.839, 85.082]
  MoveL 724 to (0, -31.52, 4.31) mm, rotated rx 8.11 ry 0 rz 180 deg; joints [17.668, -57.72, 107.959, -157.493, 52.453, 83.941]
  MoveL 725 to (0, -30.93, 4.24) mm, rotated rx 4.93 ry 0 rz 180 deg; joints [17.846, -56.754, 108.111, -157.598, 53.529, 81.163]
  MoveL 726 to (-200, -30.93, 4.24) mm, rotated rx 4.93 ry 0 rz 180 deg; joints [20.651, -66.203, 124.021, -155.996, 60.106, 82.416]
  MoveL 727 to (-200, -30.33, 4.21) mm, rotated rx 1.75 ry 0 rz 180 deg; joints [20.805, -65.019, 124.191, -156.132, 61.376, 79.778]
  MoveL 728 to (0, -30.33, 4.21) mm, rotated rx 1.75 ry 0 rz 180 deg; joints [17.982, -55.775, 108.263, -157.747, 54.607, 78.414]
  MoveL 729 to (0, -29.73, 4.2) mm, rotated rx 0 ry 0 rz 180 deg; joints [18.038, -55.221, 108.349, -157.85, 55.212, 76.925]
  MoveL 730 to (-200, -29.73, 4.2) mm, rotated rx 0 ry 0 rz 180 deg; joints [20.868, -64.349, 124.286, -156.227, 62.089, 78.35]
  MoveL 731 to (-200, -29.13, 4.2) mm, rotated rx 0 ry 0 rz 180 deg; joints [20.868, -64.315, 124.292, -156.236, 62.127, 78.368]
  MoveL 732 to (0, -29.13, 4.2) mm, rotated rx 0 ry 0 rz 180 deg; joints [18.038, -55.193, 108.355, -157.859, 55.244, 76.94]
  MoveL 733 to (0, -28.53, 4.2) mm, rotated rx 0 ry 0 rz 180 deg; joints [18.038, -55.165, 108.361, -157.868, 55.275, 76.956]
  MoveL 734 to (-200, -28.53, 4.2) mm, rotated rx 0 ry 0 rz 180 deg; joints [20.868, -64.281, 124.299, -156.245, 62.164, 78.387]
  MoveL 735 to (-200, -27.93, 4.2) mm, rotated rx 0 ry 0 rz 180 deg; joints [20.868, -64.247, 124.306, -156.253, 62.202, 78.405]
  MoveL 736 to (0, -27.93, 4.2) mm, rotated rx 0 ry 0 rz 180 deg; joints [18.038, -55.137, 108.368, -157.877, 55.307, 76.972]
  MoveL 737 to (0, -27.33, 4.2) mm, rotated rx 0 ry 0 rz 180 deg; joints [18.038, -55.109, 108.374, -157.886, 55.339, 76.987]
  MoveL 738 to (-200, -27.33, 4.2) mm, rotated rx 0 ry 0 rz 180 deg; joints [20.868, -64.213, 124.313, -156.262, 62.239, 78.424]
  MoveL 739 to (-200, -26.73, 4.2) mm, rotated rx 0 ry 0 rz 180 deg; joints [20.868, -64.179, 124.32, -156.271, 62.276, 78.443]
  MoveL 740 to (0, -26.73, 4.2) mm, rotated rx 0 ry 0 rz 180 deg; joints [18.038, -55.081, 108.38, -157.894, 55.371, 77.003]
  MoveL 741 to (0, -26.13, 4.2) mm, rotated rx 0 ry 0 rz 180 deg; joints [18.038, -55.053, 108.386, -157.903, 55.402, 77.019]
  MoveL 742 to (-200, -26.13, 4.2) mm, rotated rx 0 ry 0 rz 180 deg; joints [20.868, -64.145, 124.326, -156.279, 62.313, 78.461]
  MoveL 743 to (-200, -25.53, 4.2) mm, rotated rx 0 ry 0 rz 180 deg; joints [20.868, -64.111, 124.333, -156.288, 62.351, 78.48]
  MoveL 744 to (0, -25.53, 4.2) mm, rotated rx 0 ry 0 rz 180 deg; joints [18.038, -55.025, 108.392, -157.912, 55.434, 77.034]
  MoveL 745 to (0, -24.93, 4.2) mm, rotated rx 0 ry 0 rz 180 deg; joints [18.038, -54.997, 108.398, -157.921, 55.466, 77.05]
  MoveL 746 to (-200, -24.93, 4.2) mm, rotated rx 0 ry 0 rz 180 deg; joints [20.868, -64.076, 124.34, -156.296, 62.388, 78.498]
  MoveL 747 to (-200, -24.33, 4.2) mm, rotated rx 0 ry 0 rz 180 deg; joints [20.868, -64.042, 124.346, -156.305, 62.425, 78.517]
  MoveL 748 to (0, -24.33, 4.2) mm, rotated rx 0 ry 0 rz 180 deg; joints [18.038, -54.969, 108.405, -157.93, 55.497, 77.065]
  MoveL 749 to (0, -23.73, 4.2) mm, rotated rx 0 ry 0 rz 180 deg; joints [18.038, -54.941, 108.411, -157.939, 55.529, 77.081]
  MoveL 750 to (-200, -23.73, 4.2) mm, rotated rx 0 ry 0 rz 180 deg; joints [20.868, -64.008, 124.353, -156.314, 62.463, 78.535]
  MoveL 751 to (-200, -23.13, 4.2) mm, rotated rx 0 ry 0 rz 180 deg; joints [20.868, -63.974, 124.359, -156.322, 62.5, 78.553]
  MoveL 752 to (0, -23.13, 4.2) mm, rotated rx 0 ry 0 rz 180 deg; joints [18.038, -54.913, 108.417, -157.948, 55.561, 77.097]
  MoveL 753 to (0, -22.53, 4.2) mm, rotated rx 0 ry 0 rz 180 deg; joints [18.038, -54.884, 108.423, -157.956, 55.592, 77.112]
  MoveL 754 to (-200, -22.53, 4.2) mm, rotated rx 0 ry 0 rz 180 deg; joints [20.868, -63.94, 124.366, -156.331, 62.537, 78.572]
  MoveL 755 to (-200, -21.93, 4.2) mm, rotated rx 0 ry 0 rz 180 deg; joints [20.868, -63.906, 124.372, -156.339, 62.575, 78.59]
  MoveL 756 to (0, -21.93, 4.2) mm, rotated rx 0 ry 0 rz 180 deg; joints [18.038, -54.856, 108.429, -157.965, 55.624, 77.128]
  MoveL 757 to (0, -21.33, 4.2) mm, rotated rx 0 ry 0 rz 180 deg; joints [18.038, -54.828, 108.435, -157.974, 55.656, 77.143]
  MoveL 758 to (-200, -21.33, 4.2) mm, rotated rx 0 ry 0 rz 180 deg; joints [20.868, -63.871, 124.379, -156.347, 62.612, 78.609]
  MoveL 759 to (-200, -20.73, 4.2) mm, rotated rx 0 ry 0 rz 180 deg; joints [20.868, -63.837, 124.385, -156.356, 62.649, 78.627]
  MoveL 760 to (0, -20.73, 4.2) mm, rotated rx 0 ry 0 rz 180 deg; joints [18.038, -54.8, 108.44, -157.983, 55.687, 77.159]
  MoveL 761 to (0, -20.13, 4.2) mm, rotated rx 0 ry 0 rz 180 deg; joints [18.038, -54.772, 108.446, -157.991, 55.719, 77.174]
  MoveL 762 to (-200, -20.13, 4.2) mm, rotated rx 0 ry 0 rz 180 deg; joints [20.868, -63.803, 124.392, -156.364, 62.686, 78.645]
  MoveL 763 to (-200, -19.53, 4.2) mm, rotated rx 0 ry 0 rz 180 deg; joints [20.868, -63.769, 124.398, -156.373, 62.724, 78.664]
  MoveL 764 to (0, -19.53, 4.2) mm, rotated rx 0 ry 0 rz 180 deg; joints [18.038, -54.743, 108.452, -158, 55.75, 77.19]
  MoveL 765 to (0, -18.93, 4.2) mm, rotated rx 0 ry 0 rz 180 deg; joints [18.038, -54.715, 108.458, -158.009, 55.782, 77.205]
  MoveL 766 to (-200, -18.93, 4.2) mm, rotated rx 0 ry 0 rz 180 deg; joints [20.868, -63.734, 124.404, -156.381, 62.761, 78.682]
  MoveL 767 to (-200, -18.33, 4.2) mm, rotated rx 0 ry 0 rz 180 deg; joints [20.868, -63.7, 124.411, -156.39, 62.798, 78.7]
  MoveL 768 to (0, -18.33, 4.2) mm, rotated rx 0 ry 0 rz 180 deg; joints [18.038, -54.687, 108.464, -158.017, 55.814, 77.22]
  MoveL 769 to (0, -17.73, 4.2) mm, rotated rx 0 ry 0 rz 180 deg; joints [18.038, -54.659, 108.47, -158.026, 55.845, 77.236]
  MoveL 770 to (-200, -17.73, 4.2) mm, rotated rx 0 ry 0 rz 180 deg; joints [20.868, -63.666, 124.417, -156.398, 62.835, 78.719]
  MoveL 771 to (-200, -17.13, 4.2) mm, rotated rx 0 ry 0 rz 180 deg; joints [20.868, -63.631, 124.423, -156.406, 62.873, 78.737]
  MoveL 772 to (0, -17.13, 4.2) mm, rotated rx 0 ry 0 rz 180 deg; joints [18.038, -54.63, 108.475, -158.035, 55.877, 77.251]
  MoveL 773 to (0, -16.53, 4.2) mm, rotated rx 0 ry 0 rz 180 deg; joints [18.038, -54.602, 108.481, -158.043, 55.908, 77.267]
  MoveL 774 to (-200, -16.53, 4.2) mm, rotated rx 0 ry 0 rz 180 deg; joints [20.868, -63.597, 124.429, -156.415, 62.91, 78.755]
  MoveL 775 to (-200, -15.93, 4.2) mm, rotated rx 0 ry 0 rz 180 deg; joints [20.868, -63.562, 124.435, -156.423, 62.947, 78.773]
  MoveL 776 to (0, -15.93, 4.2) mm, rotated rx 0 ry 0 rz 180 deg; joints [18.038, -54.574, 108.487, -158.052, 55.94, 77.282]
  MoveL 777 to (0, -15.33, 4.2) mm, rotated rx 0 ry 0 rz 180 deg; joints [18.038, -54.545, 108.492, -158.06, 55.971, 77.297]
  MoveL 778 to (-200, -15.33, 4.2) mm, rotated rx 0 ry 0 rz 180 deg; joints [20.868, -63.528, 124.442, -156.431, 62.984, 78.792]
  MoveL 779 to (-200, -14.73, 4.2) mm, rotated rx 0 ry 0 rz 180 deg; joints [20.868, -63.493, 124.448, -156.439, 63.021, 78.81]
  MoveL 780 to (0, -14.73, 4.2) mm, rotated rx 0 ry 0 rz 180 deg; joints [18.038, -54.517, 108.498, -158.069, 56.003, 77.313]
  MoveL 781 to (0, -14.13, 4.2) mm, rotated rx 0 ry 0 rz 180 deg; joints [18.038, -54.489, 108.504, -158.078, 56.034, 77.328]
  MoveL 782 to (-200, -14.13, 4.2) mm, rotated rx 0 ry 0 rz 180 deg; joints [20.868, -63.459, 124.454, -156.448, 63.059, 78.828]
  MoveL 783 to (-200, -13.53, 4.2) mm, rotated rx 0 ry 0 rz 180 deg; joints [20.868, -63.424, 124.46, -156.456, 63.096, 78.846]
  MoveL 784 to (0, -13.53, 4.2) mm, rotated rx 0 ry 0 rz 180 deg; joints [18.038, -54.46, 108.509, -158.086, 56.066, 77.343]
  MoveL 785 to (0, -12.93, 4.2) mm, rotated rx 0 ry 0 rz 180 deg; joints [18.038, -54.432, 108.515, -158.095, 56.097, 77.358]
  MoveL 786 to (-200, -12.93, 4.2) mm, rotated rx 0 ry 0 rz 180 deg; joints [20.868, -63.39, 124.466, -156.464, 63.133, 78.864]
  MoveL 787 to (-200, -12.33, 4.2) mm, rotated rx 0 ry 0 rz 180 deg; joints [20.868, -63.355, 124.472, -156.472, 63.17, 78.882]
  MoveL 788 to (0, -12.33, 4.2) mm, rotated rx 0 ry 0 rz 180 deg; joints [18.038, -54.403, 108.52, -158.103, 56.129, 77.374]
  MoveL 789 to (0, -11.73, 4.2) mm, rotated rx 0 ry 0 rz 180 deg; joints [18.038, -54.375, 108.526, -158.112, 56.16, 77.389]
  MoveL 790 to (-200, -11.73, 4.2) mm, rotated rx 0 ry 0 rz 180 deg; joints [20.868, -63.321, 124.478, -156.48, 63.207, 78.901]
  MoveL 791 to (-200, -11.13, 4.2) mm, rotated rx 0 ry 0 rz 180 deg; joints [20.868, -63.286, 124.484, -156.489, 63.244, 78.919]
  MoveL 792 to (0, -11.13, 4.2) mm, rotated rx 0 ry 0 rz 180 deg; joints [18.038, -54.346, 108.531, -158.12, 56.192, 77.404]
  MoveL 793 to (0, -10.53, 4.2) mm, rotated rx 0 ry 0 rz 180 deg; joints [18.038, -54.318, 108.537, -158.129, 56.223, 77.419]
  MoveL 794 to (-200, -10.53, 4.2) mm, rotated rx 0 ry 0 rz 180 deg; joints [20.868, -63.251, 124.49, -156.497, 63.282, 78.937]
  MoveL 795 to (-200, -9.93, 4.2) mm, rotated rx 0 ry 0 rz 180 deg; joints [20.868, -63.217, 124.495, -156.505, 63.319, 78.955]
  MoveL 796 to (0, -9.93, 4.2) mm, rotated rx 0 ry 0 rz 180 deg; joints [18.038, -54.289, 108.542, -158.137, 56.255, 77.435]
  MoveL 797 to (0, -9.33, 4.2) mm, rotated rx 0 ry 0 rz 180 deg; joints [18.038, -54.261, 108.547, -158.145, 56.286, 77.45]
  MoveL 798 to (-200, -9.33, 4.2) mm, rotated rx 0 ry 0 rz 180 deg; joints [20.868, -63.182, 124.501, -156.513, 63.356, 78.973]
  MoveL 799 to (-200, -8.73, 4.2) mm, rotated rx 0 ry 0 rz 180 deg; joints [20.868, -63.148, 124.507, -156.521, 63.393, 78.991]
  MoveL 800 to (0, -8.73, 4.2) mm, rotated rx 0 ry 0 rz 180 deg; joints [18.038, -54.232, 108.553, -158.154, 56.318, 77.465]
  MoveL 801 to (0, -8.13, 4.2) mm, rotated rx 0 ry 0 rz 180 deg; joints [18.038, -54.204, 108.558, -158.162, 56.349, 77.48]
  MoveL 802 to (-200, -8.13, 4.2) mm, rotated rx 0 ry 0 rz 180 deg; joints [20.868, -63.113, 124.513, -156.529, 63.43, 79.009]
  MoveL 803 to (-200, -7.53, 4.2) mm, rotated rx 0 ry 0 rz 180 deg; joints [20.868, -63.078, 124.519, -156.537, 63.467, 79.027]
  MoveL 804 to (0, -7.53, 4.2) mm, rotated rx 0 ry 0 rz 180 deg; joints [18.038, -54.175, 108.563, -158.171, 56.381, 77.495]
  MoveL 805 to (0, -6.93, 4.2) mm, rotated rx 0 ry 0 rz 180 deg; joints [18.038, -54.147, 108.568, -158.179, 56.412, 77.51]
  MoveL 806 to (-200, -6.93, 4.2) mm, rotated rx 0 ry 0 rz 180 deg; joints [20.868, -63.043, 124.524, -156.545, 63.504, 79.045]
  MoveL 807 to (-200, -6.33, 4.2) mm, rotated rx 0 ry 0 rz 180 deg; joints [20.868, -63.009, 124.53, -156.553, 63.541, 79.063]
  MoveL 808 to (0, -6.33, 4.2) mm, rotated rx 0 ry 0 rz 180 deg; joints [18.038, -54.118, 108.574, -158.187, 56.443, 77.525]
  MoveL 809 to (0, -5.73, 4.2) mm, rotated rx 0 ry 0 rz 180 deg; joints [18.038, -54.089, 108.579, -158.196, 56.475, 77.54]
  MoveL 810 to (-200, -5.73, 4.2) mm, rotated rx 0 ry 0 rz 180 deg; joints [20.868, -62.974, 124.536, -156.561, 63.578, 79.081]
  MoveL 811 to (-200, -5.13, 4.2) mm, rotated rx 0 ry 0 rz 180 deg; joints [20.868, -62.939, 124.541, -156.569, 63.615, 79.099]
  MoveL 812 to (0, -5.13, 4.2) mm, rotated rx 0 ry 0 rz 180 deg; joints [18.038, -54.061, 108.584, -158.204, 56.506, 77.555]
  MoveL 813 to (0, -4.53, 4.2) mm, rotated rx 0 ry 0 rz 180 deg; joints [18.038, -54.032, 108.589, -158.212, 56.538, 77.57]
  MoveL 814 to (-200, -4.53, 4.2) mm, rotated rx 0 ry 0 rz 180 deg; joints [20.868, -62.904, 124.547, -156.577, 63.653, 79.117]
  MoveL 815 to (-200, -3.93, 4.2) mm, rotated rx 0 ry 0 rz 180 deg; joints [20.868, -62.869, 124.552, -156.585, 63.69, 79.135]
  MoveL 816 to (0, -3.93, 4.2) mm, rotated rx 0 ry 0 rz 180 deg; joints [18.038, -54.003, 108.594, -158.22, 56.569, 77.586]
  MoveL 817 to (0, -3.33, 4.2) mm, rotated rx 0 ry 0 rz 180 deg; joints [18.038, -53.975, 108.599, -158.229, 56.6, 77.601]
  MoveL 818 to (-200, -3.33, 4.2) mm, rotated rx 0 ry 0 rz 180 deg; joints [20.868, -62.834, 124.558, -156.593, 63.727, 79.153]
  MoveL 819 to (-200, -2.73, 4.2) mm, rotated rx 0 ry 0 rz 180 deg; joints [20.868, -62.799, 124.563, -156.601, 63.764, 79.17]
  MoveL 820 to (0, -2.73, 4.2) mm, rotated rx 0 ry 0 rz 180 deg; joints [18.038, -53.946, 108.604, -158.237, 56.632, 77.616]
  MoveL 821 to (0, -2.13, 4.2) mm, rotated rx 0 ry 0 rz 180 deg; joints [18.038, -53.917, 108.609, -158.245, 56.663, 77.631]
  MoveL 822 to (-200, -2.13, 4.2) mm, rotated rx 0 ry 0 rz 180 deg; joints [20.868, -62.765, 124.569, -156.609, 63.801, 79.188]
  MoveL 823 to (-200, -1.53, 4.2) mm, rotated rx 0 ry 0 rz 180 deg; joints [20.868, -62.73, 124.574, -156.617, 63.838, 79.206]
  MoveL 824 to (0, -1.53, 4.2) mm, rotated rx 0 ry 0 rz 180 deg; joints [18.038, -53.888, 108.614, -158.253, 56.694, 77.645]
  MoveL 825 to (0, -0.93, 4.2) mm, rotated rx 0 ry 0 rz 180 deg; joints [18.038, -53.86, 108.619, -158.262, 56.726, 77.66]
  MoveL 826 to (-200, -0.93, 4.2) mm, rotated rx 0 ry 0 rz 180 deg; joints [20.868, -62.695, 124.579, -156.625, 63.875, 79.224]
  MoveL 827 to (-200, -0.33, 4.2) mm, rotated rx 0 ry 0 rz 180 deg; joints [20.868, -62.66, 124.585, -156.632, 63.912, 79.242]
  MoveL 828 to (0, -0.33, 4.2) mm, rotated rx 0 ry 0 rz 180 deg; joints [18.038, -53.831, 108.624, -158.27, 56.757, 77.675]
  MoveL 829 to (0, 0, 4.2) mm, rotated rx 0 ry 0 rz 180 deg; joints [18.038, -53.815, 108.627, -158.274, 56.774, 77.684]
  MoveL 830 to (-200, 0, 4.2) mm, rotated rx 0 ry 0 rz 180 deg; joints [20.868, -62.64, 124.588, -156.637, 63.932, 79.252]
  MoveL 831 to (-200, 0, 3.8) mm, rotated rx 0 ry 0 rz 180 deg; joints [20.885, -62.634, 124.576, -156.617, 63.931, 79.241]
  MoveL 832 to (0, 0, 3.8) mm, rotated rx 0 ry 0 rz 180 deg; joints [18.053, -53.809, 108.616, -158.255, 56.773, 77.672]
  MoveL 833 to (0, -0.6, 3.8) mm, rotated rx 0 ry 0 rz 180 deg; joints [18.053, -53.838, 108.611, -158.247, 56.741, 77.657]
  MoveL 834 to (-200, -0.6, 3.8) mm, rotated rx 0 ry 0 rz 180 deg; joints [20.885, -62.669, 124.571, -156.609, 63.894, 79.223]
  MoveL 835 to (-200, -1.2, 3.8) mm, rotated rx 0 ry 0 rz 180 deg; joints [20.885, -62.704, 124.566, -156.601, 63.857, 79.206]
  MoveL 836 to (0, -1.2, 3.8) mm, rotated rx 0 ry 0 rz 180 deg; joints [18.053, -53.867, 108.606, -158.239, 56.71, 77.642]
  MoveL 837 to (0, -1.8, 3.8) mm, rotated rx 0 ry 0 rz 180 deg; joints [18.053, -53.895, 108.601, -158.231, 56.679, 77.627]
  MoveL 838 to (-200, -1.8, 3.8) mm, rotated rx 0 ry 0 rz 180 deg; joints [20.885, -62.739, 124.56, -156.594, 63.82, 79.188]
  MoveL 839 to (-200, -2.4, 3.8) mm, rotated rx 0 ry 0 rz 180 deg; joints [20.885, -62.774, 124.555, -156.586, 63.783, 79.17]
  MoveL 840 to (0, -2.4, 3.8) mm, rotated rx 0 ry 0 rz 180 deg; joints [18.053, -53.924, 108.596, -158.223, 56.647, 77.612]
  MoveL 841 to (0, -3, 3.8) mm, rotated rx 0 ry 0 rz 180 deg; joints [18.053, -53.953, 108.591, -158.214, 56.616, 77.597]
  MoveL 842 to (-200, -3, 3.8) mm, rotated rx 0 ry 0 rz 180 deg; joints [20.885, -62.809, 124.549, -156.578, 63.746, 79.152]
  MoveL 843 to (-200, -3.6, 3.8) mm, rotated rx 0 ry 0 rz 180 deg; joints [20.885, -62.844, 124.544, -156.57, 63.709, 79.134]
  MoveL 844 to (0, -3.6, 3.8) mm, rotated rx 0 ry 0 rz 180 deg; joints [18.053, -53.981, 108.586, -158.206, 56.585, 77.582]
  MoveL 845 to (0, -4.2, 3.8) mm, rotated rx 0 ry 0 rz 180 deg; joints [18.053, -54.01, 108.581, -158.198, 56.553, 77.567]
  MoveL 846 to (-200, -4.2, 3.8) mm, rotated rx 0 ry 0 rz 180 deg; joints [20.885, -62.878, 124.538, -156.562, 63.672, 79.116]
  MoveL 847 to (-200, -4.8, 3.8) mm, rotated rx 0 ry 0 rz 180 deg; joints [20.885, -62.913, 124.533, -156.554, 63.635, 79.098]
  MoveL 848 to (0, -4.8, 3.8) mm, rotated rx 0 ry 0 rz 180 deg; joints [18.053, -54.039, 108.576, -158.19, 56.522, 77.552]
  MoveL 849 to (0, -5.4, 3.8) mm, rotated rx 0 ry 0 rz 180 deg; joints [18.053, -54.068, 108.571, -158.181, 56.491, 77.537]
  MoveL 850 to (-200, -5.4, 3.8) mm, rotated rx 0 ry 0 rz 180 deg; joints [20.885, -62.948, 124.527, -156.546, 63.597, 79.08]
  MoveL 851 to (-200, -6, 3.8) mm, rotated rx 0 ry 0 rz 180 deg; joints [20.885, -62.983, 124.522, -156.538, 63.56, 79.062]
  MoveL 852 to (0, -6, 3.8) mm, rotated rx 0 ry 0 rz 180 deg; joints [18.053, -54.096, 108.565, -158.173, 56.459, 77.522]
  MoveL 853 to (0, -6.6, 3.8) mm, rotated rx 0 ry 0 rz 180 deg; joints [18.053, -54.125, 108.56, -158.165, 56.428, 77.506]
  MoveL 854 to (-200, -6.6, 3.8) mm, rotated rx 0 ry 0 rz 180 deg; joints [20.885, -63.018, 124.516, -156.53, 63.523, 79.044]
  MoveL 855 to (-200, -7.2, 3.8) mm, rotated rx 0 ry 0 rz 180 deg; joints [20.885, -63.052, 124.51, -156.522, 63.486, 79.026]
  MoveL 856 to (0, -7.2, 3.8) mm, rotated rx 0 ry 0 rz 180 deg; joints [18.053, -54.153, 108.555, -158.156, 56.396, 77.491]
  MoveL 857 to (0, -7.8, 3.8) mm, rotated rx 0 ry 0 rz 180 deg; joints [18.053, -54.182, 108.55, -158.148, 56.365, 77.476]
  MoveL 858 to (-200, -7.8, 3.8) mm, rotated rx 0 ry 0 rz 180 deg; joints [20.885, -63.087, 124.504, -156.514, 63.449, 79.008]
  MoveL 859 to (-200, -8.4, 3.8) mm, rotated rx 0 ry 0 rz 180 deg; joints [20.885, -63.122, 124.499, -156.506, 63.412, 78.99]
  MoveL 860 to (0, -8.4, 3.8) mm, rotated rx 0 ry 0 rz 180 deg; joints [18.053, -54.211, 108.544, -158.139, 56.334, 77.461]
  MoveL 861 to (0, -9, 3.8) mm, rotated rx 0 ry 0 rz 180 deg; joints [18.053, -54.239, 108.539, -158.131, 56.302, 77.446]
  MoveL 862 to (-200, -9, 3.8) mm, rotated rx 0 ry 0 rz 180 deg; joints [20.885, -63.157, 124.493, -156.498, 63.375, 78.972]
  MoveL 863 to (-200, -9.6, 3.8) mm, rotated rx 0 ry 0 rz 180 deg; joints [20.885, -63.191, 124.487, -156.49, 63.338, 78.954]
  MoveL 864 to (0, -9.6, 3.8) mm, rotated rx 0 ry 0 rz 180 deg; joints [18.053, -54.268, 108.534, -158.123, 56.271, 77.431]
  MoveL 865 to (0, -10.2, 3.8) mm, rotated rx 0 ry 0 rz 180 deg; joints [18.053, -54.296, 108.528, -158.114, 56.239, 77.416]
  MoveL 866 to (-200, -10.2, 3.8) mm, rotated rx 0 ry 0 rz 180 deg; joints [20.885, -63.226, 124.481, -156.481, 63.301, 78.936]
  MoveL 867 to (-200, -10.8, 3.8) mm, rotated rx 0 ry 0 rz 180 deg; joints [20.885, -63.261, 124.475, -156.473, 63.264, 78.918]
  MoveL 868 to (0, -10.8, 3.8) mm, rotated rx 0 ry 0 rz 180 deg; joints [18.053, -54.325, 108.523, -158.106, 56.208, 77.4]
  MoveL 869 to (0, -11.4, 3.8) mm, rotated rx 0 ry 0 rz 180 deg; joints [18.053, -54.353, 108.518, -158.097, 56.176, 77.385]
  MoveL 870 to (-200, -11.4, 3.8) mm, rotated rx 0 ry 0 rz 180 deg; joints [20.885, -63.295, 124.47, -156.465, 63.226, 78.9]
  MoveL 871 to (-200, -12, 3.8) mm, rotated rx 0 ry 0 rz 180 deg; joints [20.885, -63.33, 124.464, -156.457, 63.189, 78.882]
  MoveL 872 to (0, -12, 3.8) mm, rotated rx 0 ry 0 rz 180 deg; joints [18.053, -54.382, 108.512, -158.089, 56.145, 77.37]
  MoveL 873 to (0, -12.6, 3.8) mm, rotated rx 0 ry 0 rz 180 deg; joints [18.053, -54.41, 108.507, -158.08, 56.113, 77.355]
  MoveL 874 to (-200, -12.6, 3.8) mm, rotated rx 0 ry 0 rz 180 deg; joints [20.885, -63.364, 124.458, -156.449, 63.152, 78.864]
  MoveL 875 to (-200, -13.2, 3.8) mm, rotated rx 0 ry 0 rz 180 deg; joints [20.885, -63.399, 124.452, -156.441, 63.115, 78.845]
  MoveL 876 to (0, -13.2, 3.8) mm, rotated rx 0 ry 0 rz 180 deg; joints [18.053, -54.439, 108.501, -158.072, 56.082, 77.339]
  MoveL 877 to (0, -13.8, 3.8) mm, rotated rx 0 ry 0 rz 180 deg; joints [18.053, -54.467, 108.496, -158.063, 56.05, 77.324]
  MoveL 878 to (-200, -13.8, 3.8) mm, rotated rx 0 ry 0 rz 180 deg; joints [20.885, -63.433, 124.446, -156.432, 63.078, 78.827]
  MoveL 879 to (-200, -14.4, 3.8) mm, rotated rx 0 ry 0 rz 180 deg; joints [20.885, -63.468, 124.44, -156.424, 63.041, 78.809]
  MoveL 880 to (0, -14.4, 3.8) mm, rotated rx 0 ry 0 rz 180 deg; joints [18.053, -54.495, 108.49, -158.055, 56.019, 77.309]
  MoveL 881 to (0, -15, 3.8) mm, rotated rx 0 ry 0 rz 180 deg; joints [18.053, -54.524, 108.484, -158.046, 55.987, 77.293]
  MoveL 882 to (-200, -15, 3.8) mm, rotated rx 0 ry 0 rz 180 deg; joints [20.885, -63.502, 124.434, -156.416, 63.003, 78.791]
  MoveL 883 to (-200, -15.6, 3.8) mm, rotated rx 0 ry 0 rz 180 deg; joints [20.885, -63.537, 124.427, -156.408, 62.966, 78.773]
  MoveL 884 to (0, -15.6, 3.8) mm, rotated rx 0 ry 0 rz 180 deg; joints [18.053, -54.552, 108.479, -158.038, 55.956, 77.278]
  MoveL 885 to (0, -16.2, 3.8) mm, rotated rx 0 ry 0 rz 180 deg; joints [18.053, -54.58, 108.473, -158.029, 55.924, 77.263]
  MoveL 886 to (-200, -16.2, 3.8) mm, rotated rx 0 ry 0 rz 180 deg; joints [20.885, -63.571, 124.421, -156.399, 62.929, 78.754]
  MoveL 887 to (-200, -16.8, 3.8) mm, rotated rx 0 ry 0 rz 180 deg; joints [20.885, -63.606, 124.415, -156.391, 62.892, 78.736]
  MoveL 888 to (0, -16.8, 3.8) mm, rotated rx 0 ry 0 rz 180 deg; joints [18.053, -54.609, 108.467, -158.02, 55.893, 77.247]
  MoveL 889 to (0, -17.4, 3.8) mm, rotated rx 0 ry 0 rz 180 deg; joints [18.053, -54.637, 108.462, -158.012, 55.861, 77.232]
  MoveL 890 to (-200, -17.4, 3.8) mm, rotated rx 0 ry 0 rz 180 deg; joints [20.885, -63.64, 124.409, -156.383, 62.855, 78.718]
  MoveL 891 to (-200, -18, 3.8) mm, rotated rx 0 ry 0 rz 180 deg; joints [20.885, -63.674, 124.403, -156.374, 62.817, 78.7]
  MoveL 892 to (0, -18, 3.8) mm, rotated rx 0 ry 0 rz 180 deg; joints [18.053, -54.665, 108.456, -158.003, 55.83, 77.217]
  MoveL 893 to (0, -18.6, 3.8) mm, rotated rx 0 ry 0 rz 180 deg; joints [18.053, -54.694, 108.45, -157.994, 55.798, 77.201]
  MoveL 894 to (-200, -18.6, 3.8) mm, rotated rx 0 ry 0 rz 180 deg; joints [20.885, -63.709, 124.396, -156.366, 62.78, 78.681]
  MoveL 895 to (-200, -19.2, 3.8) mm, rotated rx 0 ry 0 rz 180 deg; joints [20.885, -63.743, 124.39, -156.358, 62.743, 78.663]
  MoveL 896 to (0, -19.2, 3.8) mm, rotated rx 0 ry 0 rz 180 deg; joints [18.053, -54.722, 108.444, -157.986, 55.766, 77.186]
  MoveL 897 to (0, -19.8, 3.8) mm, rotated rx 0 ry 0 rz 180 deg; joints [18.053, -54.75, 108.438, -157.977, 55.735, 77.17]
  MoveL 898 to (-200, -19.8, 3.8) mm, rotated rx 0 ry 0 rz 180 deg; joints [20.885, -63.777, 124.384, -156.349, 62.706, 78.645]
  MoveL 899 to (-200, -20.4, 3.8) mm, rotated rx 0 ry 0 rz 180 deg; joints [20.885, -63.812, 124.377, -156.341, 62.669, 78.626]
  MoveL 900 to (0, -20.4, 3.8) mm, rotated rx 0 ry 0 rz 180 deg; joints [18.053, -54.778, 108.433, -157.968, 55.703, 77.155]
  MoveL 901 to (0, -21, 3.8) mm, rotated rx 0 ry 0 rz 180 deg; joints [18.053, -54.807, 108.427, -157.96, 55.672, 77.139]
  MoveL 902 to (-200, -21, 3.8) mm, rotated rx 0 ry 0 rz 180 deg; joints [20.885, -63.846, 124.371, -156.332, 62.631, 78.608]
  MoveL 903 to (-200, -21.6, 3.8) mm, rotated rx 0 ry 0 rz 180 deg; joints [20.885, -63.88, 124.364, -156.324, 62.594, 78.59]
  MoveL 904 to (0, -21.6, 3.8) mm, rotated rx 0 ry 0 rz 180 deg; joints [18.053, -54.835, 108.421, -157.951, 55.64, 77.124]
  MoveL 905 to (0, -22.2, 3.8) mm, rotated rx 0 ry 0 rz 180 deg; joints [18.053, -54.863, 108.415, -157.942, 55.608, 77.108]
  MoveL 906 to (-200, -22.2, 3.8) mm, rotated rx 0 ry 0 rz 180 deg; joints [20.885, -63.914, 124.358, -156.315, 62.557, 78.571]
  MoveL 907 to (-200, -22.8, 3.8) mm, rotated rx 0 ry 0 rz 180 deg; joints [20.885, -63.949, 124.351, -156.307, 62.519, 78.553]
  MoveL 908 to (0, -22.8, 3.8) mm, rotated rx 0 ry 0 rz 180 deg; joints [18.053, -54.891, 108.409, -157.933, 55.577, 77.093]
  MoveL 909 to (0, -23.4, 3.8) mm, rotated rx 0 ry 0 rz 180 deg; joints [18.053, -54.919, 108.403, -157.924, 55.545, 77.077]
  MoveL 910 to (-200, -23.4, 3.8) mm, rotated rx 0 ry 0 rz 180 deg; joints [20.885, -63.983, 124.345, -156.298, 62.482, 78.534]
  MoveL 911 to (-200, -24, 3.8) mm, rotated rx 0 ry 0 rz 180 deg; joints [20.885, -64.017, 124.338, -156.29, 62.445, 78.516]
  MoveL 912 to (0, -24, 3.8) mm, rotated rx 0 ry 0 rz 180 deg; joints [18.053, -54.947, 108.397, -157.916, 55.513, 77.062]
  MoveL 913 to (0, -24.6, 3.8) mm, rotated rx 0 ry 0 rz 180 deg; joints [18.053, -54.975, 108.391, -157.907, 55.482, 77.046]
  MoveL 914 to (-200, -24.6, 3.8) mm, rotated rx 0 ry 0 rz 180 deg; joints [20.885, -64.051, 124.332, -156.281, 62.408, 78.497]
  MoveL 915 to (-200, -25.2, 3.8) mm, rotated rx 0 ry 0 rz 180 deg; joints [20.885, -64.085, 124.325, -156.273, 62.37, 78.479]
  MoveL 916 to (0, -25.2, 3.8) mm, rotated rx 0 ry 0 rz 180 deg; joints [18.053, -55.003, 108.385, -157.898, 55.45, 77.03]
  MoveL 917 to (0, -25.8, 3.8) mm, rotated rx 0 ry 0 rz 180 deg; joints [18.053, -55.031, 108.378, -157.889, 55.418, 77.015]
  MoveL 918 to (-200, -25.8, 3.8) mm, rotated rx 0 ry 0 rz 180 deg; joints [20.885, -64.119, 124.319, -156.264, 62.333, 78.46]
  MoveL 919 to (-200, -26.4, 3.8) mm, rotated rx 0 ry 0 rz 180 deg; joints [20.885, -64.153, 124.312, -156.255, 62.296, 78.442]
  MoveL 920 to (0, -26.4, 3.8) mm, rotated rx 0 ry 0 rz 180 deg; joints [18.053, -55.059, 108.372, -157.88, 55.387, 76.999]
  MoveL 921 to (0, -27, 3.8) mm, rotated rx 0 ry 0 rz 180 deg; joints [18.053, -55.087, 108.366, -157.871, 55.355, 76.984]
  MoveL 922 to (-200, -27, 3.8) mm, rotated rx 0 ry 0 rz 180 deg; joints [20.885, -64.187, 124.305, -156.247, 62.258, 78.423]
  MoveL 923 to (-200, -27.6, 3.8) mm, rotated rx 0 ry 0 rz 180 deg; joints [20.885, -64.221, 124.298, -156.238, 62.221, 78.405]
  MoveL 924 to (0, -27.6, 3.8) mm, rotated rx 0 ry 0 rz 180 deg; joints [18.053, -55.115, 108.36, -157.862, 55.323, 76.968]
  MoveL 925 to (0, -28.2, 3.8) mm, rotated rx 0 ry 0 rz 180 deg; joints [18.053, -55.143, 108.354, -157.853, 55.292, 76.952]
  MoveL 926 to (-200, -28.2, 3.8) mm, rotated rx 0 ry 0 rz 180 deg; joints [20.885, -64.255, 124.292, -156.23, 62.184, 78.386]
  MoveL 927 to (-200, -28.8, 3.8) mm, rotated rx 0 ry 0 rz 180 deg; joints [20.885, -64.289, 124.285, -156.221, 62.146, 78.367]
  MoveL 928 to (0, -28.8, 3.8) mm, rotated rx 0 ry 0 rz 180 deg; joints [18.053, -55.171, 108.347, -157.844, 55.26, 76.936]
  MoveL 929 to (0, -29.4, 3.8) mm, rotated rx 0 ry 0 rz 180 deg; joints [18.053, -55.199, 108.341, -157.836, 55.228, 76.921]
  MoveL 930 to (-200, -29.4, 3.8) mm, rotated rx 0 ry 0 rz 180 deg; joints [20.885, -64.323, 124.278, -156.212, 62.109, 78.349]
  MoveL 931 to (-200, -30, 3.8) mm, rotated rx 0 ry 0 rz 180 deg; joints [20.885, -64.357, 124.271, -156.203, 62.072, 78.33]
  MoveL 932 to (0, -30, 3.8) mm, rotated rx 0 ry 0 rz 180 deg; joints [18.053, -55.227, 108.335, -157.827, 55.197, 76.905]
  MoveL 933 to (0, -30.6, 3.82) mm, rotated rx 3.07 ry 0 rz 180 deg; joints [17.946, -56.178, 108.189, -157.66, 54.157, 79.539]
  MoveL 934 to (-200, -30.6, 3.82) mm, rotated rx 3.07 ry 0 rz 180 deg; joints [20.764, -65.507, 124.109, -156.05, 60.846, 80.859]
  MoveL 935 to (-200, -31.2, 3.86) mm, rotated rx 6.14 ry 0 rz 180 deg; joints [20.597, -66.644, 123.944, -155.934, 59.622, 83.412]
  MoveL 936 to (0, -31.2, 3.86) mm, rotated rx 6.14 ry 0 rz 180 deg; joints [17.798, -57.118, 108.042, -157.533, 53.117, 82.2]
  MoveL 937 to (0, -31.79, 3.94) mm, rotated rx 9.21 ry 0 rz 180 deg; joints [17.612, -58.045, 107.895, -157.447, 52.079, 84.89]
  MoveL 938 to (-200, -31.79, 3.94) mm, rotated rx 9.21 ry 0 rz 180 deg; joints [20.386, -67.764, 123.778, -155.859, 58.4, 85.993]
  MoveL 939 to (-200, -32.38, 4.06) mm, rotated rx 12.28 ry 0 rz 180 deg; joints [20.129, -68.864, 123.61, -155.827, 57.184, 88.606]
  MoveL 940 to (0, -32.38, 4.06) mm, rotated rx 12.28 ry 0 rz 180 deg; joints [17.385, -58.957, 107.748, -157.404, 51.045, 87.615]
  MoveL 941 to (0, -32.96, 4.2) mm, rotated rx 15.35 ry 0 rz 180 deg; joints [17.12, -59.852, 107.602, -157.407, 50.016, 90.377]
  MoveL 942 to (-200, -32.96, 4.2) mm, rotated rx 15.35 ry 0 rz 180 deg; joints [19.829, -69.943, 123.443, -155.84, 55.975, 91.257]
  MoveL 943 to (-200, -33.54, 4.37) mm, rotated rx 18.42 ry 0 rz 180 deg; joints [19.484, -70.998, 123.277, -155.902, 54.776, 93.951]
  MoveL 944 to (0, -33.54, 4.37) mm, rotated rx 18.42 ry 0 rz 180 deg; joints [16.816, -60.728, 107.458, -157.459, 48.996, 93.183]
  MoveL 945 to (0, -34.1, 4.58) mm, rotated rx 21.49 ry 0 rz 180 deg; joints [16.474, -61.581, 107.317, -157.562, 47.986, 96.036]
  MoveL 946 to (-200, -34.1, 4.58) mm, rotated rx 21.49 ry 0 rz 180 deg; joints [19.095, -72.025, 123.113, -156.015, 53.589, 96.692]
  MoveL 947 to (-200, -34.65, 4.81) mm, rotated rx 24.55 ry 0 rz 180 deg; joints [18.664, -73.024, 122.951, -156.183, 52.417, 99.487]
  MoveL 948 to (0, -34.65, 4.81) mm, rotated rx 24.55 ry 0 rz 180 deg; joints [16.095, -62.412, 107.18, -157.72, 46.989, 98.94]
  MoveL 949 to (0, -35.19, 5.08) mm, rotated rx 27.63 ry 0 rz 180 deg; joints [15.679, -63.217, 107.047, -157.936, 46.008, 101.902]
  MoveL 950 to (-200, -35.19, 5.08) mm, rotated rx 27.63 ry 0 rz 180 deg; joints [18.19, -73.993, 122.794, -156.409, 51.262, 102.341]
  MoveL 951 to (-200, -35.72, 5.37) mm, rotated rx 30.69 ry 0 rz 180 deg; joints [17.675, -74.928, 122.642, -156.697, 50.129, 105.258]
  MoveL 952 to (0, -35.72, 5.37) mm, rotated rx 30.69 ry 0 rz 180 deg; joints [15.227, -63.995, 106.919, -158.214, 45.045, 104.924]
  MoveL 953 to (0, -36.23, 5.69) mm, rotated rx 33.76 ry 0 rz 180 deg; joints [14.74, -64.745, 106.798, -158.556, 44.103, 108.013]
  MoveL 954 to (-200, -36.23, 5.69) mm, rotated rx 33.76 ry 0 rz 180 deg; joints [17.118, -75.827, 122.496, -157.051, 49.018, 108.245]
  MoveL 955 to (-200, -36.71, 6.04) mm, rotated rx 36.83 ry 0 rz 180 deg; joints [16.522, -76.69, 122.358, -157.476, 47.936, 111.306]
  MoveL 956 to (0, -36.71, 6.04) mm, rotated rx 36.83 ry 0 rz 180 deg; joints [14.219, -65.463, 106.684, -158.967, 43.187, 111.171]
  MoveL 957 to (0, -37.19, 6.41) mm, rotated rx 39.9 ry 0 rz 180 deg; joints [13.666, -66.149, 106.578, -159.448, 42.298, 114.403]
  MoveL 958 to (-200, -37.19, 6.41) mm, rotated rx 39.9 ry 0 rz 180 deg; joints [15.888, -77.513, 122.228, -157.974, 46.884, 114.446]
  MoveL 959 to (-200, -37.63, 6.8) mm, rotated rx 42.97 ry 0 rz 180 deg; joints [15.216, -78.296, 122.108, -158.551, 45.867, 117.672]
  MoveL 960 to (0, -37.63, 6.8) mm, rotated rx 42.97 ry 0 rz 180 deg; joints [13.08, -66.801, 106.482, -160.005, 41.44, 117.714]
  MoveL 961 to (0, -38.06, 7.23) mm, rotated rx 46.04 ry 0 rz 180 deg; joints [12.464, -67.418, 106.396, -160.638, 40.618, 121.106]
  MoveL 962 to (-200, -38.06, 7.23) mm, rotated rx 46.04 ry 0 rz 180 deg; joints [14.508, -79.036, 121.998, -159.209, 44.89, 120.985]
  MoveL 963 to (-200, -38.47, 7.67) mm, rotated rx 49.11 ry 0 rz 180 deg; joints [13.765, -79.732, 121.901, -159.951, 43.955, 124.392]
  MoveL 964 to (0, -38.47, 7.67) mm, rotated rx 49.11 ry 0 rz 180 deg; joints [11.82, -67.997, 106.32, -161.351, 39.835, 124.582]
  MoveL 965 to (0, -38.85, 8.13) mm, rotated rx 52.18 ry 0 rz 180 deg; joints [11.148, -68.539, 106.256, -162.145, 39.094, 128.144]
  MoveL 966 to (-200, -38.85, 8.13) mm, rotated rx 52.18 ry 0 rz 180 deg; joints [12.991, -80.382, 121.816, -160.781, 43.07, 127.892]
  MoveL 967 to (-200, -39.2, 8.62) mm, rotated rx 55.25 ry 0 rz 180 deg; joints [12.185, -80.984, 121.745, -161.699, 42.237, 131.491]
  MoveL 968 to (0, -39.2, 8.62) mm, rotated rx 55.25 ry 0 rz 180 deg; joints [10.451, -69.041, 106.205, -163.021, 38.401, 131.793]
  MoveL 969 to (0, -39.53, 9.12) mm, rotated rx 58.32 ry 0 rz 180 deg; joints [9.731, -69.502, 106.168, -163.977, 37.759, 135.527]
  MoveL 970 to (-200, -39.53, 9.12) mm, rotated rx 58.32 ry 0 rz 180 deg; joints [11.351, -81.538, 121.689, -162.707, 41.463, 135.186]
  MoveL 971 to (-200, -39.83, 9.64) mm, rotated rx 61.39 ry 0 rz 180 deg; joints [10.491, -82.041, 121.649, -163.803, 40.752, 138.978]
  MoveL 972 to (0, -39.83, 9.64) mm, rotated rx 61.39 ry 0 rz 180 deg; joints [8.989, -69.921, 106.144, -165.014, 37.173, 139.347]
  MoveL 973 to (0, -40.1, 10.17) mm, rotated rx 64.46 ry 0 rz 180 deg; joints [8.228, -70.297, 106.134, -166.128, 36.646, 143.25]
  MoveL 974 to (-200, -40.1, 10.17) mm, rotated rx 64.46 ry 0 rz 180 deg; joints [9.607, -82.493, 121.625, -164.986, 40.11, 142.866]
  MoveL 975 to (-200, -40.35, 10.72) mm, rotated rx 67.53 ry 0 rz 180 deg; joints [8.703, -82.892, 121.618, -166.251, 39.541, 146.842]
  MoveL 976 to (0, -40.35, 10.72) mm, rotated rx 67.53 ry 0 rz 180 deg; joints [7.449, -70.629, 106.14, -167.314, 36.183, 147.229]
  MoveL 977 to (0, -40.56, 11.28) mm, rotated rx 70.6 ry 0 rz 180 deg; joints [6.656, -70.916, 106.161, -168.568, 35.788, 151.281]
  MoveL 978 to (-200, -40.56, 11.28) mm, rotated rx 70.6 ry 0 rz 180 deg; joints [7.779, -83.238, 121.628, -167.593, 39.051, 150.902]
  MoveL 979 to (-200, -40.75, 11.85) mm, rotated rx 73.67 ry 0 rz 180 deg; joints [6.841, -83.529, 121.657, -169.004, 38.645, 155.037]
  MoveL 980 to (0, -40.75, 11.85) mm, rotated rx 73.67 ry 0 rz 180 deg; joints [5.851, -71.158, 106.198, -169.88, 35.464, 155.395]
  MoveL 981 to (0, -40.9, 12.43) mm, rotated rx 76.73 ry 0 rz 180 deg; joints [5.036, -71.353, 106.251, -171.243, 35.214, 159.562]
  MoveL 982 to (-200, -40.9, 12.43) mm, rotated rx 76.73 ry 0 rz 180 deg; joints [5.89, -83.764, 121.703, -170.475, 38.325, 159.236]
  MoveL 983 to (-200, -41.02, 13.02) mm, rotated rx 79.81 ry 0 rz 180 deg; joints [4.93, -83.944, 121.769, -171.994, 38.097, 163.489]
  MoveL 984 to (0, -41.02, 13.02) mm, rotated rx 79.81 ry 0 rz 180 deg; joints [4.214, -71.501, 106.319, -172.647, 35.04, 163.774]
  MoveL 985 to (0, -41.11, 13.61) mm, rotated rx 82.87 ry 0 rz 180 deg; joints [3.387, -71.602, 106.404, -174.079, 34.946, 168.015]
  MoveL 986 to (-200, -41.11, 13.61) mm, rotated rx 82.87 ry 0 rz 180 deg; joints [3.964, -84.066, 121.852, -173.548, 37.963, 167.779]
  MoveL 987 to (-200, -41.17, 14.21) mm, rotated rx 85.94 ry 0 rz 180 deg; joints [2.995, -84.131, 121.954, -175.124, 37.924, 172.094]
  MoveL 988 to (0, -41.17, 14.21) mm, rotated rx 85.94 ry 0 rz 180 deg; joints [2.559, -71.655, 106.504, -175.528, 34.931, 172.275]
  MoveL 989 to (0, -41.2, 14.81) mm, rotated rx 89.01 ry 0 rz 180 deg; joints [1.731, -71.659, 106.619, -176.98, 34.998, 176.538]
  MoveL 990 to (-200, -41.2, 14.81) mm, rotated rx 89.01 ry 0 rz 180 deg; joints [2.027, -84.137, 122.074, -176.706, 37.982, 176.415]
  MoveL 991 to (-200, -41.2, 15.41) mm, rotated rx 90 ry 0 rz 180 deg; joints [1.696, -84.128, 122.117, -177.245, 38.021, 177.829]
  MoveL 992 to (0, -41.2, 15.41) mm, rotated rx 90 ry 0 rz 180 deg; joints [1.449, -71.651, 106.661, -177.475, 35.036, 177.932]
  MoveL 993 to (0, -41.2, 16.01) mm, rotated rx 90 ry 0 rz 180 deg; joints [1.424, -71.652, 106.662, -177.519, 35.035, 177.968]
  MoveL 994 to (-200, -41.2, 16.01) mm, rotated rx 90 ry 0 rz 180 deg; joints [1.667, -84.129, 122.118, -177.293, 38.02, 177.867]
  MoveL 995 to (-200, -41.2, 16.61) mm, rotated rx 90 ry 0 rz 180 deg; joints [1.638, -84.13, 122.12, -177.341, 38.019, 177.904]
  MoveL 996 to (0, -41.2, 16.61) mm, rotated rx 90 ry 0 rz 180 deg; joints [1.399, -71.653, 106.663, -177.563, 35.035, 178.004]
  MoveL 997 to (0, -41.2, 17.21) mm, rotated rx 90 ry 0 rz 180 deg; joints [1.374, -71.654, 106.664, -177.606, 35.034, 178.04]
  MoveL 998 to (-200, -41.2, 17.21) mm, rotated rx 90 ry 0 rz 180 deg; joints [1.608, -84.131, 122.121, -177.388, 38.018, 177.942]
  MoveL 999 to (-200, -41.2, 17.81) mm, rotated rx 90 ry 0 rz 180 deg; joints [1.579, -84.132, 122.122, -177.436, 38.017, 177.979]
  MoveL 1000 to (0, -41.2, 17.81) mm, rotated rx 90 ry 0 rz 180 deg; joints [1.349, -71.654, 106.665, -177.65, 35.034, 178.075]
  MoveL 1001 to (0, -41.2, 18.41) mm, rotated rx 90 ry 0 rz 180 deg; joints [1.324, -71.655, 106.667, -177.693, 35.033, 178.111]
  MoveL 1002 to (-200, -41.2, 18.41) mm, rotated rx 90 ry 0 rz 180 deg; joints [1.55, -84.134, 122.123, -177.483, 38.017, 178.017]
  MoveL 1003 to (-200, -41.2, 19.01) mm, rotated rx 90 ry 0 rz 180 deg; joints [1.52, -84.135, 122.124, -177.531, 38.016, 178.054]
  MoveL 1004 to (0, -41.2, 19.01) mm, rotated rx 90 ry 0 rz 180 deg; joints [1.299, -71.656, 106.668, -177.737, 35.033, 178.147]
  MoveL 1005 to (0, -41.2, 19.61) mm, rotated rx 90 ry 0 rz 180 deg; joints [1.274, -71.657, 106.669, -177.781, 35.032, 178.182]
  MoveL 1006 to (-200, -41.2, 19.61) mm, rotated rx 90 ry 0 rz 180 deg; joints [1.491, -84.136, 122.126, -177.578, 38.015, 178.092]
  MoveL 1007 to (-200, -41.2, 20.21) mm, rotated rx 90 ry 0 rz 180 deg; joints [1.462, -84.137, 122.127, -177.626, 38.014, 178.129]
  MoveL 1008 to (0, -41.2, 20.21) mm, rotated rx 90 ry 0 rz 180 deg; joints [1.249, -71.658, 106.67, -177.824, 35.032, 178.218]
  MoveL 1009 to (0, -41.2, 20.81) mm, rotated rx 90 ry 0 rz 180 deg; joints [1.224, -71.659, 106.671, -177.868, 35.031, 178.254]
  MoveL 1010 to (-200, -41.2, 20.81) mm, rotated rx 90 ry 0 rz 180 deg; joints [1.432, -84.138, 122.128, -177.674, 38.013, 178.167]
  MoveL 1011 to (-200, -41.2, 21.41) mm, rotated rx 90 ry 0 rz 180 deg; joints [1.403, -84.138, 122.129, -177.721, 38.012, 178.204]
  MoveL 1012 to (0, -41.2, 21.41) mm, rotated rx 90 ry 0 rz 180 deg; joints [1.199, -71.659, 106.672, -177.912, 35.031, 178.29]
  MoveL 1013 to (0, -41.2, 22.01) mm, rotated rx 90 ry 0 rz 180 deg; joints [1.174, -71.66, 106.673, -177.955, 35.03, 178.325]
  MoveL 1014 to (-200, -41.2, 22.01) mm, rotated rx 90 ry 0 rz 180 deg; joints [1.374, -84.139, 122.13, -177.769, 38.012, 178.242]
  MoveL 1015 to (-200, -41.2, 22.61) mm, rotated rx 90 ry 0 rz 180 deg; joints [1.344, -84.14, 122.131, -177.816, 38.011, 178.279]
  MoveL 1016 to (0, -41.2, 22.61) mm, rotated rx 90 ry 0 rz 180 deg; joints [1.149, -71.661, 106.674, -177.999, 35.03, 178.361]
  MoveL 1017 to (0, -41.2, 23.21) mm, rotated rx 90 ry 0 rz 180 deg; joints [1.124, -71.662, 106.675, -178.042, 35.029, 178.397]
  MoveL 1018 to (-200, -41.2, 23.21) mm, rotated rx 90 ry 0 rz 180 deg; joints [1.315, -84.141, 122.132, -177.864, 38.01, 178.317]
  MoveL 1019 to (-200, -41.2, 23.81) mm, rotated rx 90 ry 0 rz 180 deg; joints [1.286, -84.142, 122.133, -177.912, 38.009, 178.354]
  MoveL 1020 to (0, -41.2, 23.81) mm, rotated rx 90 ry 0 rz 180 deg; joints [1.098, -71.662, 106.676, -178.086, 35.029, 178.433]
  MoveL 1021 to (0, -41.2, 24.41) mm, rotated rx 90 ry 0 rz 180 deg; joints [1.073, -71.663, 106.677, -178.13, 35.028, 178.468]
  MoveL 1022 to (-200, -41.2, 24.41) mm, rotated rx 90 ry 0 rz 180 deg; joints [1.257, -84.143, 122.134, -177.959, 38.009, 178.392]
  MoveL 1023 to (-200, -41.2, 25.01) mm, rotated rx 90 ry 0 rz 180 deg; joints [1.227, -84.144, 122.135, -178.007, 38.008, 178.429]
  MoveL 1024 to (0, -41.2, 25.01) mm, rotated rx 90 ry 0 rz 180 deg; joints [1.048, -71.664, 106.678, -178.173, 35.028, 178.504]
  MoveL 1025 to (0, -41.2, 25.61) mm, rotated rx 90 ry 0 rz 180 deg; joints [1.023, -71.664, 106.679, -178.217, 35.028, 178.54]
  MoveL 1026 to (-200, -41.2, 25.61) mm, rotated rx 90 ry 0 rz 180 deg; joints [1.198, -84.145, 122.136, -178.054, 38.007, 178.467]
  MoveL 1027 to (-200, -41.2, 26.21) mm, rotated rx 90 ry 0 rz 180 deg; joints [1.169, -84.145, 122.137, -178.102, 38.006, 178.504]
  MoveL 1028 to (0, -41.2, 26.21) mm, rotated rx 90 ry 0 rz 180 deg; joints [0.998, -71.665, 106.68, -178.261, 35.027, 178.575]
  MoveL 1029 to (0, -41.2, 26.81) mm, rotated rx 90 ry 0 rz 180 deg; joints [0.973, -71.666, 106.681, -178.304, 35.027, 178.611]
  MoveL 1030 to (-200, -41.2, 26.81) mm, rotated rx 90 ry 0 rz 180 deg; joints [1.139, -84.146, 122.137, -178.15, 38.006, 178.542]
  MoveL 1031 to (-200, -41.2, 27.41) mm, rotated rx 90 ry 0 rz 180 deg; joints [1.11, -84.147, 122.138, -178.197, 38.005, 178.579]
  MoveL 1032 to (0, -41.2, 27.41) mm, rotated rx 90 ry 0 rz 180 deg; joints [0.948, -71.666, 106.682, -178.348, 35.026, 178.647]
  MoveL 1033 to (0, -41.2, 28.01) mm, rotated rx 90 ry 0 rz 180 deg; joints [0.923, -71.667, 106.682, -178.392, 35.026, 178.683]
  MoveL 1034 to (-200, -41.2, 28.01) mm, rotated rx 90 ry 0 rz 180 deg; joints [1.081, -84.148, 122.139, -178.245, 38.004, 178.617]
  MoveL 1035 to (-200, -41.2, 28.61) mm, rotated rx 90 ry 0 rz 180 deg; joints [1.051, -84.148, 122.14, -178.292, 38.004, 178.654]
  MoveL 1036 to (0, -41.2, 28.61) mm, rotated rx 90 ry 0 rz 180 deg; joints [0.898, -71.668, 106.683, -178.435, 35.026, 178.718]
  MoveL 1037 to (0, -41.2, 29.21) mm, rotated rx 90 ry 0 rz 180 deg; joints [0.873, -71.668, 106.684, -178.479, 35.025, 178.754]
  MoveL 1038 to (-200, -41.2, 29.21) mm, rotated rx 90 ry 0 rz 180 deg; joints [1.022, -84.149, 122.141, -178.34, 38.003, 178.692]
  MoveL 1039 to (-200, -41.2, 29.81) mm, rotated rx 90 ry 0 rz 180 deg; joints [0.993, -84.15, 122.141, -178.388, 38.003, 178.729]
  MoveL 1040 to (0, -41.2, 29.81) mm, rotated rx 90 ry 0 rz 180 deg; joints [0.848, -71.669, 106.685, -178.522, 35.025, 178.79]
  MoveL 1041 to (0, -41.2, 30.41) mm, rotated rx 90 ry 0 rz 180 deg; joints [0.823, -71.669, 106.685, -178.566, 35.025, 178.826]
  MoveL 1042 to (-200, -41.2, 30.41) mm, rotated rx 90 ry 0 rz 180 deg; joints [0.963, -84.15, 122.142, -178.435, 38.002, 178.767]
  MoveL 1043 to (-200, -41.2, 31.01) mm, rotated rx 90 ry 0 rz 180 deg; joints [0.934, -84.151, 122.143, -178.483, 38.002, 178.804]
  MoveL 1044 to (0, -41.2, 31.01) mm, rotated rx 90 ry 0 rz 180 deg; joints [0.798, -71.67, 106.686, -178.61, 35.024, 178.861]
  MoveL 1045 to (0, -41.2, 31.61) mm, rotated rx 90 ry 0 rz 180 deg; joints [0.773, -71.67, 106.687, -178.653, 35.024, 178.897]
  MoveL 1046 to (-200, -41.2, 31.61) mm, rotated rx 90 ry 0 rz 180 deg; joints [0.905, -84.152, 122.144, -178.531, 38.001, 178.842]
  MoveL 1047 to (-200, -41.2, 32.21) mm, rotated rx 90 ry 0 rz 180 deg; joints [0.875, -84.152, 122.144, -178.578, 38.001, 178.879]
  MoveL 1048 to (0, -41.2, 32.21) mm, rotated rx 90 ry 0 rz 180 deg; joints [0.748, -71.671, 106.687, -178.697, 35.024, 178.933]
  MoveL 1049 to (0, -41.2, 32.81) mm, rotated rx 90 ry 0 rz 180 deg; joints [0.723, -71.671, 106.688, -178.741, 35.023, 178.969]
  MoveL 1050 to (-200, -41.2, 32.81) mm, rotated rx 90 ry 0 rz 180 deg; joints [0.846, -84.153, 122.145, -178.626, 38, 178.917]
  MoveL 1051 to (-200, -41.2, 33.41) mm, rotated rx 90 ry 0 rz 180 deg; joints [0.817, -84.153, 122.146, -178.673, 38, 178.955]
  MoveL 1052 to (0, -41.2, 33.41) mm, rotated rx 90 ry 0 rz 180 deg; joints [0.698, -71.672, 106.689, -178.784, 35.023, 179.004]
  MoveL 1053 to (0, -41.2, 34.01) mm, rotated rx 90 ry 0 rz 180 deg; joints [0.673, -71.672, 106.689, -178.828, 35.023, 179.04]
  MoveL 1054 to (-200, -41.2, 34.01) mm, rotated rx 90 ry 0 rz 180 deg; joints [0.787, -84.154, 122.146, -178.721, 37.999, 178.992]
  MoveL 1055 to (-200, -41.2, 34.61) mm, rotated rx 90 ry 0 rz 180 deg; joints [0.758, -84.154, 122.147, -178.769, 37.999, 179.03]
  MoveL 1056 to (0, -41.2, 34.61) mm, rotated rx 90 ry 0 rz 180 deg; joints [0.648, -71.672, 106.69, -178.872, 35.023, 179.076]
  MoveL 1057 to (0, -41.2, 35.21) mm, rotated rx 90 ry 0 rz 180 deg; joints [0.622, -71.673, 106.69, -178.915, 35.022, 179.112]
  MoveL 1058 to (-200, -41.2, 35.21) mm, rotated rx 90 ry 0 rz 180 deg; joints [0.729, -84.155, 122.147, -178.816, 37.998, 179.067]
  MoveL 1059 to (-200, -41.2, 35.81) mm, rotated rx 90 ry 0 rz 180 deg; joints [0.699, -84.155, 122.148, -178.864, 37.998, 179.105]
  MoveL 1060 to (0, -41.2, 35.81) mm, rotated rx 90 ry 0 rz 180 deg; joints [0.597, -71.673, 106.691, -178.959, 35.022, 179.147]
  MoveL 1061 to (0, -41.2, 36.41) mm, rotated rx 90 ry 0 rz 180 deg; joints [0.572, -71.674, 106.691, -179.003, 35.022, 179.183]
  MoveL 1062 to (-200, -41.2, 36.41) mm, rotated rx 90 ry 0 rz 180 deg; joints [0.67, -84.156, 122.148, -178.912, 37.997, 179.142]
  MoveL 1063 to (-200, -41.2, 37.01) mm, rotated rx 90 ry 0 rz 180 deg; joints [0.641, -84.156, 122.149, -178.959, 37.997, 179.18]
  MoveL 1064 to (0, -41.2, 37.01) mm, rotated rx 90 ry 0 rz 180 deg; joints [0.547, -71.674, 106.692, -179.046, 35.022, 179.219]
  MoveL 1065 to (0, -41.2, 37.61) mm, rotated rx 90 ry 0 rz 180 deg; joints [0.522, -71.674, 106.692, -179.09, 35.021, 179.255]
  MoveL 1066 to (-200, -41.2, 37.61) mm, rotated rx 90 ry 0 rz 180 deg; joints [0.611, -84.157, 122.149, -179.007, 37.997, 179.217]
  MoveL 1067 to (-200, -41.2, 38.21) mm, rotated rx 90 ry 0 rz 180 deg; joints [0.582, -84.157, 122.15, -179.054, 37.996, 179.255]
  MoveL 1068 to (0, -41.2, 38.21) mm, rotated rx 90 ry 0 rz 180 deg; joints [0.497, -71.675, 106.693, -179.134, 35.021, 179.29]
  MoveL 1069 to (0, -41.2, 38.81) mm, rotated rx 90 ry 0 rz 180 deg; joints [0.472, -71.675, 106.693, -179.177, 35.021, 179.326]
  MoveL 1070 to (-200, -41.2, 38.81) mm, rotated rx 90 ry 0 rz 180 deg; joints [0.553, -84.158, 122.15, -179.102, 37.996, 179.292]
  MoveL 1071 to (-200, -41.2, 39.41) mm, rotated rx 90 ry 0 rz 180 deg; joints [0.523, -84.158, 122.151, -179.15, 37.996, 179.33]
  MoveL 1072 to (0, -41.2, 39.41) mm, rotated rx 90 ry 0 rz 180 deg; joints [0.447, -71.675, 106.694, -179.221, 35.021, 179.362]
  MoveL 1073 to (0, -41.2, 40.01) mm, rotated rx 90 ry 0 rz 180 deg; joints [0.422, -71.676, 106.694, -179.265, 35.021, 179.398]
  MoveL 1074 to (-200, -41.2, 40.01) mm, rotated rx 90 ry 0 rz 180 deg; joints [0.494, -84.158, 122.151, -179.197, 37.995, 179.368]
  MoveL 1075 to (-200, -41.2, 40.61) mm, rotated rx 90 ry 0 rz 180 deg; joints [0.465, -84.159, 122.151, -179.245, 37.995, 179.405]
  MoveL 1076 to (0, -41.2, 40.61) mm, rotated rx 90 ry 0 rz 180 deg; joints [0.397, -71.676, 106.694, -179.308, 35.021, 179.433]
  MoveL 1077 to (0, -41.2, 41.21) mm, rotated rx 90 ry 0 rz 180 deg; joints [0.372, -71.676, 106.695, -179.352, 35.02, 179.469]
  MoveL 1078 to (-200, -41.2, 41.21) mm, rotated rx 90 ry 0 rz 180 deg; joints [0.435, -84.159, 122.152, -179.293, 37.995, 179.443]
  MoveL 1079 to (-200, -41.2, 41.81) mm, rotated rx 90 ry 0 rz 180 deg; joints [0.406, -84.159, 122.152, -179.34, 37.995, 179.48]
  MoveL 1080 to (0, -41.2, 41.81) mm, rotated rx 90 ry 0 rz 180 deg; joints [0.347, -71.676, 106.695, -179.396, 35.02, 179.505]
  MoveL 1081 to (0, -41.2, 42.41) mm, rotated rx 90 ry 0 rz 180 deg; joints [0.322, -71.677, 106.695, -179.439, 35.02, 179.541]
  MoveL 1082 to (-200, -41.2, 42.41) mm, rotated rx 90 ry 0 rz 180 deg; joints [0.377, -84.159, 122.152, -179.388, 37.994, 179.518]
  MoveL 1083 to (-200, -41.2, 43.01) mm, rotated rx 90 ry 0 rz 180 deg; joints [0.347, -84.16, 122.153, -179.436, 37.994, 179.555]
  MoveL 1084 to (0, -41.2, 43.01) mm, rotated rx 90 ry 0 rz 180 deg; joints [0.297, -71.677, 106.696, -179.483, 35.02, 179.576]
  MoveL 1085 to (0, -41.2, 43.61) mm, rotated rx 90 ry 0 rz 180 deg; joints [0.272, -71.677, 106.696, -179.527, 35.02, 179.612]
  MoveL 1086 to (-200, -41.2, 43.61) mm, rotated rx 90 ry 0 rz 180 deg; joints [0.318, -84.16, 122.153, -179.483, 37.994, 179.593]
  MoveL 1087 to (-200, -41.2, 44.21) mm, rotated rx 90 ry 0 rz 180 deg; joints [0.289, -84.16, 122.153, -179.531, 37.994, 179.63]
  MoveL 1088 to (0, -41.2, 44.21) mm, rotated rx 90 ry 0 rz 180 deg; joints [0.247, -71.677, 106.696, -179.57, 35.02, 179.648]
  MoveL 1089 to (0, -41.2, 44.81) mm, rotated rx 90 ry 0 rz 180 deg; joints [0.222, -71.677, 106.696, -179.614, 35.02, 179.684]
  MoveL 1090 to (-200, -41.2, 44.81) mm, rotated rx 90 ry 0 rz 180 deg; joints [0.259, -84.16, 122.153, -179.579, 37.994, 179.668]
  MoveL 1091 to (-200, -41.19, 45.41) mm, rotated rx 92.08 ry 0 rz 180 deg; joints [-0.404, -84.097, 122.224, 179.346, 38.129, -177.402]
  MoveL 1092 to (0, -41.19, 45.41) mm, rotated rx 92.08 ry 0 rz 180 deg; joints [-0.345, -71.624, 106.762, 179.4, 35.139, -177.427]
  MoveL 1093 to (0, -41.16, 46.01) mm, rotated rx 95.15 ry 0 rz 180 deg; joints [-1.162, -71.506, 106.872, 177.992, 35.383, -173.211]
  MoveL 1094 to (-200, -41.16, 46.01) mm, rotated rx 95.15 ry 0 rz 180 deg; joints [-1.361, -83.955, 122.343, 177.81, 38.408, -173.131]
  MoveL 1095 to (-200, -41.09, 46.6) mm, rotated rx 98.22 ry 0 rz 180 deg; joints [-2.306, -83.756, 122.478, 176.317, 38.781, -168.907]
  MoveL 1096 to (0, -41.09, 46.6) mm, rotated rx 98.22 ry 0 rz 180 deg; joints [-1.97, -71.339, 106.995, 176.623, 35.704, -169.036]
  MoveL 1097 to (0, -40.98, 47.19) mm, rotated rx 101.29 ry 0 rz 180 deg; joints [-2.765, -71.124, 107.133, 175.303, 36.1, -164.911]
  MoveL 1098 to (-200, -40.98, 47.19) mm, rotated rx 101.29 ry 0 rz 180 deg; joints [-3.236, -83.498, 122.63, 174.88, 39.244, -164.74]
  MoveL 1099 to (-200, -40.85, 47.78) mm, rotated rx 104.36 ry 0 rz 180 deg; joints [-4.149, -83.183, 122.797, 173.509, 39.795, -160.644]
  MoveL 1100 to (0, -40.85, 47.78) mm, rotated rx 104.36 ry 0 rz 180 deg; joints [-3.546, -70.862, 107.283, 174.041, 36.569, -160.848]
  MoveL 1101 to (0, -40.69, 48.35) mm, rotated rx 107.43 ry 0 rz 180 deg; joints [-4.31, -70.553, 107.445, 172.845, 37.107, -156.853]
  MoveL 1102 to (-200, -40.69, 48.35) mm, rotated rx 107.43 ry 0 rz 180 deg; joints [-5.042, -82.812, 122.978, 172.212, 40.428, -156.626]
  MoveL 1103 to (-200, -40.49, 48.92) mm, rotated rx 110.5 ry 0 rz 180 deg; joints [-5.91, -82.384, 123.172, 170.995, 41.14, -152.695]
  MoveL 1104 to (0, -40.49, 48.92) mm, rotated rx 110.5 ry 0 rz 180 deg; joints [-5.054, -70.197, 107.618, 171.72, 37.711, -152.934]
  MoveL 1105 to (0, -40.27, 49.48) mm, rotated rx 113.57 ry 0 rz 180 deg; joints [-5.776, -69.796, 107.801, 170.671, 38.376, -149.094]
  MoveL 1106 to (-200, -40.27, 49.48) mm, rotated rx 113.57 ry 0 rz 180 deg; joints [-6.753, -81.901, 123.378, 169.864, 41.925, -148.856]
  MoveL 1107 to (-200, -40.01, 50.02) mm, rotated rx 116.64 ry 0 rz 180 deg; joints [-7.567, -81.363, 123.595, 168.82, 42.779, -145.108]
  MoveL 1108 to (0, -40.01, 50.02) mm, rotated rx 116.64 ry 0 rz 180 deg; joints [-6.474, -69.35, 107.994, 169.701, 39.098, -145.335]
  MoveL 1109 to (0, -39.73, 50.55) mm, rotated rx 119.71 ry 0 rz 180 deg; joints [-7.146, -68.86, 108.194, 168.812, 39.874, -141.661]
  MoveL 1110 to (-200, -39.73, 50.55) mm, rotated rx 119.71 ry 0 rz 180 deg; joints [-8.349, -80.772, 123.822, 167.866, 43.696, -141.457]
  MoveL 1111 to (-200, -39.42, 51.06) mm, rotated rx 122.78 ry 0 rz 180 deg; joints [-9.099, -80.129, 124.056, 167.001, 44.671, -137.9]
  MoveL 1112 to (0, -39.42, 51.06) mm, rotated rx 122.78 ry 0 rz 180 deg; joints [-7.79, -68.327, 108.4, 168.002, 40.698, -138.07]
  MoveL 1113 to (0, -39.08, 51.56) mm, rotated rx 125.85 ry 0 rz 180 deg; joints [-8.405, -67.752, 108.612, 167.273, 41.566, -134.563]
  MoveL 1114 to (-200, -39.08, 51.56) mm, rotated rx 125.85 ry 0 rz 180 deg; joints [-9.813, -79.434, 124.297, 166.223, 45.699, -134.436]
  MoveL 1115 to (-200, -38.71, 52.04) mm, rotated rx 128.92 ry 0 rz 180 deg; joints [-10.49, -78.69, 124.543, 165.53, 46.775, -131.062]
  MoveL 1116 to (0, -38.71, 52.04) mm, rotated rx 128.92 ry 0 rz 180 deg; joints [-8.988, -67.137, 108.829, 166.623, 42.476, -131.136]
  MoveL 1117 to (0, -38.33, 52.49) mm, rotated rx 131.99 ry 0 rz 180 deg; joints [-9.539, -66.482, 109.048, 166.049, 43.421, -127.787]
  MoveL 1118 to (-200, -38.33, 52.49) mm, rotated rx 131.99 ry 0 rz 180 deg; joints [-11.129, -77.897, 124.792, 164.921, 47.895, -127.775]
  MoveL 1119 to (-200, -37.91, 52.93) mm, rotated rx 135.05 ry 0 rz 180 deg; joints [-11.727, -77.059, 125.043, 164.39, 49.053, -124.57]
  MoveL 1120 to (0, -37.91, 52.93) mm, rotated rx 135.05 ry 0 rz 180 deg; joints [-10.055, -65.79, 109.268, 165.549, 44.399, -124.513]
  MoveL 1121 to (0, -37.48, 53.34) mm, rotated rx 138.12 ry 0 rz 180 deg; joints [-10.536, -65.062, 109.489, 165.121, 45.405, -121.309]
  MoveL 1122 to (-200, -37.48, 53.34) mm, rotated rx 138.12 ry 0 rz 180 deg; joints [-12.283, -76.175, 125.295, 163.935, 50.246, -121.442]
  MoveL 1123 to (-200, -37.02, 53.73) mm, rotated rx 141.19 ry 0 rz 180 deg; joints [-12.797, -75.249, 125.546, 163.552, 51.469, -118.386]
  MoveL 1124 to (0, -37.02, 53.73) mm, rotated rx 141.19 ry 0 rz 180 deg; joints [-10.98, -64.299, 109.709, 164.76, 46.436, -118.173]
  MoveL 1125 to (0, -36.54, 54.09) mm, rotated rx 144.26 ry 0 rz 180 deg; joints [-11.387, -63.503, 109.927, 164.464, 47.488, -115.097]
  MoveL 1126 to (-200, -36.54, 54.09) mm, rotated rx 144.26 ry 0 rz 180 deg; joints [-13.267, -74.282, 125.794, 163.237, 52.718, -115.397]
  MoveL 1127 to (-200, -36.05, 54.43) mm, rotated rx 147.33 ry 0 rz 180 deg; joints [-13.692, -73.276, 126.038, 162.986, 53.99, -112.469]
  MoveL 1128 to (0, -36.05, 54.43) mm, rotated rx 147.33 ry 0 rz 180 deg; joints [-11.756, -62.677, 110.142, 164.229, 48.558, -112.08]
  MoveL 1129 to (0, -35.53, 54.74) mm, rotated rx 150.4 ry 0 rz 180 deg; joints [-12.085, -61.822, 110.352, 164.053, 49.643, -109.116]
  MoveL 1130 to (-200, -35.53, 54.74) mm, rotated rx 150.4 ry 0 rz 180 deg; joints [-14.071, -72.235, 126.277, 162.795, 55.28, -109.597]
  MoveL 1131 to (-200, -35, 55.02) mm, rotated rx 153.47 ry 0 rz 180 deg; joints [-14.404, -71.159, 126.51, 162.661, 56.586, -106.774]
  MoveL 1132 to (0, -35, 55.02) mm, rotated rx 153.47 ry 0 rz 180 deg; joints [-12.374, -60.94, 110.557, 163.932, 50.739, -106.199]
  MoveL 1133 to (0, -34.46, 55.27) mm, rotated rx 156.54 ry 0 rz 180 deg; joints [-12.623, -60.035, 110.755, 163.864, 51.844, -103.326]
  MoveL 1134 to (-200, -34.46, 55.27) mm, rotated rx 156.54 ry 0 rz 180 deg; joints [-14.69, -70.053, 126.734, 162.581, 57.904, -103.996]
  MoveL 1135 to (-200, -33.9, 55.5) mm, rotated rx 159.61 ry 0 rz 180 deg; joints [-14.929, -68.919, 126.95, 162.552, 59.23, -101.255]
  MoveL 1136 to (0, -33.9, 55.5) mm, rotated rx 159.61 ry 0 rz 180 deg; joints [-12.831, -59.106, 110.945, 163.845, 52.955, -100.491]
  MoveL 1137 to (0, -33.34, 55.69) mm, rotated rx 162.68 ry 0 rz 180 deg; joints [-12.997, -58.159, 111.127, 163.873, 54.068, -97.691]
  MoveL 1138 to (-200, -33.34, 55.69) mm, rotated rx 162.68 ry 0 rz 180 deg; joints [-15.121, -67.76, 127.155, 162.571, 60.562, -98.55]
  MoveL 1139 to (-200, -32.76, 55.85) mm, rotated rx 165.75 ry 0 rz 180 deg; joints [-15.264, -66.578, 127.35, 162.635, 61.897, -95.871]
  MoveL 1140 to (0, -32.76, 55.85) mm, rotated rx 165.75 ry 0 rz 180 deg; joints [-13.122, -57.194, 111.3, 163.946, 55.182, -94.92]
  MoveL 1141 to (0, -32.17, 55.99) mm, rotated rx 168.82 ry 0 rz 180 deg; joints [-13.205, -56.215, 111.463, 164.062, 56.293, -92.177]
  MoveL 1142 to (-200, -32.17, 55.99) mm, rotated rx 168.82 ry 0 rz 180 deg; joints [-15.359, -65.377, 127.532, 162.743, 63.231, -93.217]
  MoveL 1143 to (-200, -31.58, 56.09) mm, rotated rx 171.89 ry 0 rz 180 deg; joints [-15.406, -64.161, 127.702, 162.892, 64.561, -90.581]
  MoveL 1144 to (0, -31.58, 56.09) mm, rotated rx 171.89 ry 0 rz 180 deg; joints [-13.246, -55.224, 111.616, 164.218, 57.398, -89.454]
  MoveL 1145 to (0, -30.98, 56.16) mm, rotated rx 174.96 ry 0 rz 180 deg; joints [-13.244, -54.224, 111.757, 164.413, 58.497, -86.749]
  MoveL 1146 to (-200, -30.98, 56.16) mm, rotated rx 174.96 ry 0 rz 180 deg; joints [-15.404, -62.932, 127.858, 163.081, 65.885, -87.958]
  MoveL 1147 to (-200, -30.39, 56.19) mm, rotated rx 178.03 ry 0 rz 180 deg; joints [-15.354, -61.695, 128.001, 163.308, 67.2, -85.346]
  MoveL 1148 to (0, -30.39, 56.19) mm, rotated rx 178.03 ry 0 rz 180 deg; joints [-13.201, -53.218, 111.887, 164.645, 59.586, -84.06]
  MoveL 1149 to (0, -29.79, 56.2) mm, rotated rx 180 ry 0 rz 180 deg; joints [-13.15, -52.558, 111.965, 164.815, 60.291, -82.339]
  MoveL 1150 to (-200, -29.79, 56.2) mm, rotated rx 180 ry 0 rz 180 deg; joints [-15.297, -60.882, 128.086, 163.475, 68.054, -83.673]
  MoveL 1151 to (-200, -29.19, 56.2) mm, rotated rx 180 ry 0 rz 180 deg; joints [-15.297, -60.844, 128.088, 163.48, 68.093, -83.685]
  MoveL 1152 to (0, -29.19, 56.2) mm, rotated rx 180 ry 0 rz 180 deg; joints [-13.15, -52.527, 111.967, 164.82, 60.323, -82.349]
  MoveL 1153 to (0, -28.59, 56.2) mm, rotated rx 180 ry 0 rz 180 deg; joints [-13.15, -52.496, 111.969, 164.825, 60.356, -82.359]
  MoveL 1154 to (-200, -28.59, 56.2) mm, rotated rx 180 ry 0 rz 180 deg; joints [-15.297, -60.805, 128.091, 163.485, 68.132, -83.698]
  MoveL 1155 to (-200, -27.99, 56.2) mm, rotated rx 180 ry 0 rz 180 deg; joints [-15.297, -60.767, 128.093, 163.489, 68.171, -83.71]
  MoveL 1156 to (0, -27.99, 56.2) mm, rotated rx 180 ry 0 rz 180 deg; joints [-13.15, -52.464, 111.971, 164.83, 60.388, -82.369]
  MoveL 1157 to (0, -27.39, 56.2) mm, rotated rx 180 ry 0 rz 180 deg; joints [-13.15, -52.433, 111.973, 164.835, 60.42, -82.379]
  MoveL 1158 to (-200, -27.39, 56.2) mm, rotated rx 180 ry 0 rz 180 deg; joints [-15.297, -60.728, 128.095, 163.494, 68.211, -83.723]
  MoveL 1159 to (-200, -26.79, 56.2) mm, rotated rx 180 ry 0 rz 180 deg; joints [-15.297, -60.69, 128.097, 163.499, 68.25, -83.735]
  MoveL 1160 to (0, -26.79, 56.2) mm, rotated rx 180 ry 0 rz 180 deg; joints [-13.15, -52.401, 111.975, 164.84, 60.453, -82.389]
  MoveL 1161 to (0, -26.19, 56.2) mm, rotated rx 180 ry 0 rz 180 deg; joints [-13.15, -52.37, 111.977, 164.845, 60.485, -82.399]
  MoveL 1162 to (-200, -26.19, 56.2) mm, rotated rx 180 ry 0 rz 180 deg; joints [-15.297, -60.651, 128.099, 163.503, 68.289, -83.748]
  MoveL 1163 to (-200, -25.59, 56.2) mm, rotated rx 180 ry 0 rz 180 deg; joints [-15.297, -60.612, 128.102, 163.508, 68.328, -83.76]
  MoveL 1164 to (0, -25.59, 56.2) mm, rotated rx 180 ry 0 rz 180 deg; joints [-13.15, -52.338, 111.979, 164.85, 60.517, -82.41]
  MoveL 1165 to (0, -24.99, 56.2) mm, rotated rx 180 ry 0 rz 180 deg; joints [-13.15, -52.307, 111.981, 164.855, 60.549, -82.42]
  MoveL 1166 to (-200, -24.99, 56.2) mm, rotated rx 180 ry 0 rz 180 deg; joints [-15.297, -60.574, 128.104, 163.513, 68.367, -83.773]
  MoveL 1167 to (-200, -24.39, 56.2) mm, rotated rx 180 ry 0 rz 180 deg; joints [-15.297, -60.535, 128.106, 163.517, 68.406, -83.785]
  MoveL 1168 to (0, -24.39, 56.2) mm, rotated rx 180 ry 0 rz 180 deg; joints [-13.15, -52.275, 111.983, 164.86, 60.582, -82.43]
  MoveL 1169 to (0, -23.79, 56.2) mm, rotated rx 180 ry 0 rz 180 deg; joints [-13.15, -52.244, 111.985, 164.864, 60.614, -82.44]
  MoveL 1170 to (-200, -23.79, 56.2) mm, rotated rx 180 ry 0 rz 180 deg; joints [-15.297, -60.496, 128.108, 163.522, 68.445, -83.798]
  MoveL 1171 to (-200, -23.19, 56.2) mm, rotated rx 180 ry 0 rz 180 deg; joints [-15.297, -60.458, 128.11, 163.526, 68.484, -83.81]
  MoveL 1172 to (0, -23.19, 56.2) mm, rotated rx 180 ry 0 rz 180 deg; joints [-13.15, -52.212, 111.987, 164.869, 60.646, -82.45]
  MoveL 1173 to (0, -22.59, 56.2) mm, rotated rx 180 ry 0 rz 180 deg; joints [-13.15, -52.181, 111.989, 164.874, 60.678, -82.46]
  MoveL 1174 to (-200, -22.59, 56.2) mm, rotated rx 180 ry 0 rz 180 deg; joints [-15.297, -60.419, 128.112, 163.531, 68.523, -83.822]
  MoveL 1175 to (-200, -21.99, 56.2) mm, rotated rx 180 ry 0 rz 180 deg; joints [-15.297, -60.38, 128.114, 163.535, 68.562, -83.835]
  MoveL 1176 to (0, -21.99, 56.2) mm, rotated rx 180 ry 0 rz 180 deg; joints [-13.15, -52.149, 111.99, 164.879, 60.71, -82.47]
  MoveL 1177 to (0, -21.39, 56.2) mm, rotated rx 180 ry 0 rz 180 deg; joints [-13.15, -52.118, 111.992, 164.884, 60.743, -82.479]
  MoveL 1178 to (-200, -21.39, 56.2) mm, rotated rx 180 ry 0 rz 180 deg; joints [-15.297, -60.341, 128.116, 163.54, 68.601, -83.847]
  MoveL 1179 to (-200, -20.79, 56.2) mm, rotated rx 180 ry 0 rz 180 deg; joints [-15.297, -60.303, 128.117, 163.544, 68.64, -83.86]
  MoveL 1180 to (0, -20.79, 56.2) mm, rotated rx 180 ry 0 rz 180 deg; joints [-13.15, -52.086, 111.994, 164.889, 60.775, -82.489]
  MoveL 1181 to (0, -20.19, 56.2) mm, rotated rx 180 ry 0 rz 180 deg; joints [-13.15, -52.054, 111.995, 164.894, 60.807, -82.499]
  MoveL 1182 to (-200, -20.19, 56.2) mm, rotated rx 180 ry 0 rz 180 deg; joints [-15.297, -60.264, 128.119, 163.549, 68.679, -83.872]
  MoveL 1183 to (-200, -19.59, 56.2) mm, rotated rx 180 ry 0 rz 180 deg; joints [-15.297, -60.225, 128.121, 163.553, 68.718, -83.884]
  MoveL 1184 to (0, -19.59, 56.2) mm, rotated rx 180 ry 0 rz 180 deg; joints [-13.15, -52.023, 111.997, 164.899, 60.839, -82.509]
  MoveL 1185 to (0, -18.99, 56.2) mm, rotated rx 180 ry 0 rz 180 deg; joints [-13.15, -51.991, 111.999, 164.903, 60.871, -82.519]
  MoveL 1186 to (-200, -18.99, 56.2) mm, rotated rx 180 ry 0 rz 180 deg; joints [-15.297, -60.186, 128.123, 163.558, 68.757, -83.897]
  MoveL 1187 to (-200, -18.39, 56.2) mm, rotated rx 180 ry 0 rz 180 deg; joints [-15.297, -60.147, 128.125, 163.562, 68.796, -83.909]
  MoveL 1188 to (0, -18.39, 56.2) mm, rotated rx 180 ry 0 rz 180 deg; joints [-13.15, -51.959, 112, 164.908, 60.903, -82.529]
  MoveL 1189 to (0, -17.79, 56.2) mm, rotated rx 180 ry 0 rz 180 deg; joints [-13.15, -51.928, 112.002, 164.913, 60.935, -82.539]
  MoveL 1190 to (-200, -17.79, 56.2) mm, rotated rx 180 ry 0 rz 180 deg; joints [-15.297, -60.109, 128.126, 163.567, 68.835, -83.921]
  MoveL 1191 to (-200, -17.19, 56.2) mm, rotated rx 180 ry 0 rz 180 deg; joints [-15.297, -60.07, 128.128, 163.571, 68.874, -83.934]
  MoveL 1192 to (0, -17.19, 56.2) mm, rotated rx 180 ry 0 rz 180 deg; joints [-13.15, -51.896, 112.003, 164.918, 60.967, -82.549]
  MoveL 1193 to (0, -16.59, 56.2) mm, rotated rx 180 ry 0 rz 180 deg; joints [-13.15, -51.864, 112.005, 164.923, 60.999, -82.559]
  MoveL 1194 to (-200, -16.59, 56.2) mm, rotated rx 180 ry 0 rz 180 deg; joints [-15.297, -60.031, 128.13, 163.576, 68.913, -83.946]
  MoveL 1195 to (-200, -15.99, 56.2) mm, rotated rx 180 ry 0 rz 180 deg; joints [-15.297, -59.992, 128.131, 163.58, 68.952, -83.958]
  MoveL 1196 to (0, -15.99, 56.2) mm, rotated rx 180 ry 0 rz 180 deg; joints [-13.15, -51.832, 112.006, 164.927, 61.031, -82.569]
  MoveL 1197 to (0, -15.39, 56.2) mm, rotated rx 180 ry 0 rz 180 deg; joints [-13.15, -51.801, 112.008, 164.932, 61.063, -82.579]
  MoveL 1198 to (-200, -15.39, 56.2) mm, rotated rx 180 ry 0 rz 180 deg; joints [-15.297, -59.953, 128.133, 163.584, 68.99, -83.97]
  MoveL 1199 to (-200, -14.79, 56.2) mm, rotated rx 180 ry 0 rz 180 deg; joints [-15.297, -59.914, 128.134, 163.589, 69.029, -83.983]
  MoveL 1200 to (0, -14.79, 56.2) mm, rotated rx 180 ry 0 rz 180 deg; joints [-13.15, -51.769, 112.009, 164.937, 61.095, -82.588]
  MoveL 1201 to (0, -14.19, 56.2) mm, rotated rx 180 ry 0 rz 180 deg; joints [-13.15, -51.737, 112.01, 164.942, 61.127, -82.598]
  MoveL 1202 to (-200, -14.19, 56.2) mm, rotated rx 180 ry 0 rz 180 deg; joints [-15.297, -59.875, 128.136, 163.593, 69.068, -83.995]
  MoveL 1203 to (-200, -13.59, 56.2) mm, rotated rx 180 ry 0 rz 180 deg; joints [-15.297, -59.836, 128.137, 163.598, 69.107, -84.007]
  MoveL 1204 to (0, -13.59, 56.2) mm, rotated rx 180 ry 0 rz 180 deg; joints [-13.15, -51.705, 112.012, 164.946, 61.159, -82.608]
  MoveL 1205 to (0, -12.99, 56.2) mm, rotated rx 180 ry 0 rz 180 deg; joints [-13.15, -51.674, 112.013, 164.951, 61.191, -82.618]
  MoveL 1206 to (-200, -12.99, 56.2) mm, rotated rx 180 ry 0 rz 180 deg; joints [-15.297, -59.797, 128.139, 163.602, 69.146, -84.019]
  MoveL 1207 to (-200, -12.39, 56.2) mm, rotated rx 180 ry 0 rz 180 deg; joints [-15.297, -59.758, 128.14, 163.606, 69.185, -84.032]
  MoveL 1208 to (0, -12.39, 56.2) mm, rotated rx 180 ry 0 rz 180 deg; joints [-13.15, -51.642, 112.014, 164.956, 61.223, -82.628]
  MoveL 1209 to (0, -11.79, 56.2) mm, rotated rx 180 ry 0 rz 180 deg; joints [-13.15, -51.61, 112.016, 164.961, 61.255, -82.637]
  MoveL 1210 to (-200, -11.79, 56.2) mm, rotated rx 180 ry 0 rz 180 deg; joints [-15.297, -59.719, 128.142, 163.611, 69.223, -84.044]
  MoveL 1211 to (-200, -11.19, 56.2) mm, rotated rx 180 ry 0 rz 180 deg; joints [-15.297, -59.68, 128.143, 163.615, 69.262, -84.056]
  MoveL 1212 to (0, -11.19, 56.2) mm, rotated rx 180 ry 0 rz 180 deg; joints [-13.15, -51.578, 112.017, 164.965, 61.287, -82.647]
  MoveL 1213 to (0, -10.59, 56.2) mm, rotated rx 180 ry 0 rz 180 deg; joints [-13.15, -51.546, 112.018, 164.97, 61.319, -82.657]
  MoveL 1214 to (-200, -10.59, 56.2) mm, rotated rx 180 ry 0 rz 180 deg; joints [-15.297, -59.641, 128.144, 163.619, 69.301, -84.068]
  MoveL 1215 to (-200, -9.99, 56.2) mm, rotated rx 180 ry 0 rz 180 deg; joints [-15.297, -59.602, 128.146, 163.623, 69.34, -84.08]
  MoveL 1216 to (0, -9.99, 56.2) mm, rotated rx 180 ry 0 rz 180 deg; joints [-13.15, -51.514, 112.019, 164.975, 61.351, -82.667]
  MoveL 1217 to (0, -9.39, 56.2) mm, rotated rx 180 ry 0 rz 180 deg; joints [-13.15, -51.482, 112.02, 164.979, 61.383, -82.677]
  MoveL 1218 to (-200, -9.39, 56.2) mm, rotated rx 180 ry 0 rz 180 deg; joints [-15.297, -59.563, 128.147, 163.628, 69.378, -84.093]
  MoveL 1219 to (-200, -8.79, 56.2) mm, rotated rx 180 ry 0 rz 180 deg; joints [-15.297, -59.523, 128.148, 163.632, 69.417, -84.105]
  MoveL 1220 to (0, -8.79, 56.2) mm, rotated rx 180 ry 0 rz 180 deg; joints [-13.15, -51.451, 112.021, 164.984, 61.415, -82.686]
  MoveL 1221 to (0, -8.19, 56.2) mm, rotated rx 180 ry 0 rz 180 deg; joints [-13.15, -51.419, 112.022, 164.989, 61.447, -82.696]
  MoveL 1222 to (-200, -8.19, 56.2) mm, rotated rx 180 ry 0 rz 180 deg; joints [-15.297, -59.484, 128.149, 163.636, 69.456, -84.117]
  MoveL 1223 to (-200, -7.59, 56.2) mm, rotated rx 180 ry 0 rz 180 deg; joints [-15.297, -59.445, 128.15, 163.641, 69.494, -84.129]
  MoveL 1224 to (0, -7.59, 56.2) mm, rotated rx 180 ry 0 rz 180 deg; joints [-13.15, -51.387, 112.023, 164.993, 61.479, -82.706]
  MoveL 1225 to (0, -6.99, 56.2) mm, rotated rx 180 ry 0 rz 180 deg; joints [-13.15, -51.355, 112.024, 164.998, 61.511, -82.715]
  MoveL 1226 to (-200, -6.99, 56.2) mm, rotated rx 180 ry 0 rz 180 deg; joints [-15.297, -59.406, 128.152, 163.645, 69.533, -84.141]
  MoveL 1227 to (-200, -6.39, 56.2) mm, rotated rx 180 ry 0 rz 180 deg; joints [-15.297, -59.367, 128.153, 163.649, 69.572, -84.153]
  MoveL 1228 to (0, -6.39, 56.2) mm, rotated rx 180 ry 0 rz 180 deg; joints [-13.15, -51.323, 112.025, 165.003, 61.542, -82.725]
  MoveL 1229 to (0, -5.79, 56.2) mm, rotated rx 180 ry 0 rz 180 deg; joints [-13.15, -51.291, 112.026, 165.007, 61.574, -82.735]
  MoveL 1230 to (-200, -5.79, 56.2) mm, rotated rx 180 ry 0 rz 180 deg; joints [-15.297, -59.327, 128.154, 163.653, 69.61, -84.165]
  MoveL 1231 to (-200, -5.19, 56.2) mm, rotated rx 180 ry 0 rz 180 deg; joints [-15.297, -59.288, 128.155, 163.657, 69.649, -84.177]
  MoveL 1232 to (0, -5.19, 56.2) mm, rotated rx 180 ry 0 rz 180 deg; joints [-13.15, -51.259, 112.027, 165.012, 61.606, -82.745]
  MoveL 1233 to (0, -4.59, 56.2) mm, rotated rx 180 ry 0 rz 180 deg; joints [-13.15, -51.227, 112.028, 165.016, 61.638, -82.754]
  MoveL 1234 to (-200, -4.59, 56.2) mm, rotated rx 180 ry 0 rz 180 deg; joints [-15.297, -59.249, 128.156, 163.662, 69.688, -84.189]
  MoveL 1235 to (-200, -3.99, 56.2) mm, rotated rx 180 ry 0 rz 180 deg; joints [-15.297, -59.21, 128.157, 163.666, 69.726, -84.202]
  MoveL 1236 to (0, -3.99, 56.2) mm, rotated rx 180 ry 0 rz 180 deg; joints [-13.15, -51.195, 112.029, 165.021, 61.67, -82.764]
  MoveL 1237 to (0, -3.39, 56.2) mm, rotated rx 180 ry 0 rz 180 deg; joints [-13.15, -51.163, 112.03, 165.026, 61.701, -82.773]
  MoveL 1238 to (-200, -3.39, 56.2) mm, rotated rx 180 ry 0 rz 180 deg; joints [-15.297, -59.17, 128.158, 163.67, 69.765, -84.214]
  MoveL 1239 to (-200, -2.79, 56.2) mm, rotated rx 180 ry 0 rz 180 deg; joints [-15.297, -59.131, 128.158, 163.674, 69.803, -84.226]
  MoveL 1240 to (0, -2.79, 56.2) mm, rotated rx 180 ry 0 rz 180 deg; joints [-13.15, -51.131, 112.031, 165.03, 61.733, -82.783]
  MoveL 1241 to (0, -2.19, 56.2) mm, rotated rx 180 ry 0 rz 180 deg; joints [-13.15, -51.098, 112.031, 165.035, 61.765, -82.793]
  MoveL 1242 to (-200, -2.19, 56.2) mm, rotated rx 180 ry 0 rz 180 deg; joints [-15.297, -59.092, 128.159, 163.678, 69.842, -84.238]
  MoveL 1243 to (-200, -1.59, 56.2) mm, rotated rx 180 ry 0 rz 180 deg; joints [-15.297, -59.052, 128.16, 163.682, 69.881, -84.25]
  MoveL 1244 to (0, -1.59, 56.2) mm, rotated rx 180 ry 0 rz 180 deg; joints [-13.15, -51.066, 112.032, 165.039, 61.797, -82.802]
  MoveL 1245 to (0, -0.99, 56.2) mm, rotated rx 180 ry 0 rz 180 deg; joints [-13.15, -51.034, 112.033, 165.044, 61.828, -82.812]
  MoveL 1246 to (-200, -0.99, 56.2) mm, rotated rx 180 ry 0 rz 180 deg; joints [-15.297, -59.013, 128.161, 163.687, 69.919, -84.262]
  MoveL 1247 to (-200, -0.39, 56.2) mm, rotated rx 180 ry 0 rz 180 deg; joints [-15.297, -58.974, 128.162, 163.691, 69.958, -84.274]
  MoveL 1248 to (0, -0.39, 56.2) mm, rotated rx 180 ry 0 rz 180 deg; joints [-13.15, -51.002, 112.034, 165.048, 61.86, -82.822]
  MoveL 1249 to (0, 0, 56.2) mm, rotated rx 180 ry 0 rz 180 deg; joints [-13.15, -50.981, 112.034, 165.051, 61.88, -82.828]
  MoveL 1250 to (-200, 0, 56.2) mm, rotated rx 180 ry 0 rz 180 deg; joints [-15.297, -58.948, 128.162, 163.693, 69.982, -84.281]
  MoveL 1251 to (-200, 0, 56.6) mm, rotated rx 180 ry 0 rz 180 deg; joints [-15.315, -58.944, 128.154, 163.674, 69.98, -84.274]
  MoveL 1252 to (0, 0, 56.6) mm, rotated rx 180 ry 0 rz 180 deg; joints [-13.166, -50.977, 112.026, 165.033, 61.878, -82.818]
  MoveL 1253 to (0, -0.6, 56.6) mm, rotated rx 180 ry 0 rz 180 deg; joints [-13.166, -51.01, 112.025, 165.028, 61.847, -82.809]
  MoveL 1254 to (-200, -0.6, 56.6) mm, rotated rx 180 ry 0 rz 180 deg; joints [-15.315, -58.984, 128.153, 163.67, 69.942, -84.261]
  MoveL 1255 to (-200, -1.2, 56.6) mm, rotated rx 180 ry 0 rz 180 deg; joints [-15.315, -59.023, 128.152, 163.665, 69.903, -84.249]
  MoveL 1256 to (0, -1.2, 56.6) mm, rotated rx 180 ry 0 rz 180 deg; joints [-13.166, -51.042, 112.025, 165.024, 61.815, -82.799]
  MoveL 1257 to (0, -1.8, 56.6) mm, rotated rx 180 ry 0 rz 180 deg; joints [-13.166, -51.074, 112.024, 165.019, 61.783, -82.789]
  MoveL 1258 to (-200, -1.8, 56.6) mm, rotated rx 180 ry 0 rz 180 deg; joints [-15.315, -59.062, 128.151, 163.661, 69.865, -84.237]
  MoveL 1259 to (-200, -2.4, 56.6) mm, rotated rx 180 ry 0 rz 180 deg; joints [-15.315, -59.102, 128.151, 163.657, 69.826, -84.225]
  MoveL 1260 to (0, -2.4, 56.6) mm, rotated rx 180 ry 0 rz 180 deg; joints [-13.166, -51.106, 112.023, 165.015, 61.752, -82.78]
  MoveL 1261 to (0, -3, 56.6) mm, rotated rx 180 ry 0 rz 180 deg; joints [-13.166, -51.138, 112.022, 165.01, 61.72, -82.77]
  MoveL 1262 to (-200, -3, 56.6) mm, rotated rx 180 ry 0 rz 180 deg; joints [-15.315, -59.141, 128.15, 163.653, 69.787, -84.213]
  MoveL 1263 to (-200, -3.6, 56.6) mm, rotated rx 180 ry 0 rz 180 deg; joints [-15.315, -59.18, 128.149, 163.649, 69.749, -84.201]
  MoveL 1264 to (0, -3.6, 56.6) mm, rotated rx 180 ry 0 rz 180 deg; joints [-13.166, -51.17, 112.022, 165.006, 61.688, -82.76]
  MoveL 1265 to (0, -4.2, 56.6) mm, rotated rx 180 ry 0 rz 180 deg; joints [-13.166, -51.202, 112.021, 165.001, 61.656, -82.751]
  MoveL 1266 to (-200, -4.2, 56.6) mm, rotated rx 180 ry 0 rz 180 deg; joints [-15.315, -59.22, 128.148, 163.645, 69.71, -84.189]
  MoveL 1267 to (-200, -4.8, 56.6) mm, rotated rx 180 ry 0 rz 180 deg; joints [-15.315, -59.259, 128.147, 163.64, 69.672, -84.177]
  MoveL 1268 to (0, -4.8, 56.6) mm, rotated rx 180 ry 0 rz 180 deg; joints [-13.166, -51.234, 112.02, 164.996, 61.625, -82.741]
  MoveL 1269 to (0, -5.4, 56.6) mm, rotated rx 180 ry 0 rz 180 deg; joints [-13.166, -51.266, 112.019, 164.992, 61.593, -82.731]
  MoveL 1270 to (-200, -5.4, 56.6) mm, rotated rx 180 ry 0 rz 180 deg; joints [-15.315, -59.298, 128.146, 163.636, 69.633, -84.165]
  MoveL 1271 to (-200, -6, 56.6) mm, rotated rx 180 ry 0 rz 180 deg; joints [-15.315, -59.337, 128.145, 163.632, 69.594, -84.153]
  MoveL 1272 to (0, -6, 56.6) mm, rotated rx 180 ry 0 rz 180 deg; joints [-13.166, -51.298, 112.018, 164.987, 61.561, -82.722]
  MoveL 1273 to (0, -6.6, 56.6) mm, rotated rx 180 ry 0 rz 180 deg; joints [-13.166, -51.33, 112.017, 164.982, 61.529, -82.712]
  MoveL 1274 to (-200, -6.6, 56.6) mm, rotated rx 180 ry 0 rz 180 deg; joints [-15.315, -59.377, 128.144, 163.628, 69.556, -84.141]
  MoveL 1275 to (-200, -7.2, 56.6) mm, rotated rx 180 ry 0 rz 180 deg; joints [-15.315, -59.416, 128.143, 163.624, 69.517, -84.129]
  MoveL 1276 to (0, -7.2, 56.6) mm, rotated rx 180 ry 0 rz 180 deg; joints [-13.166, -51.362, 112.016, 164.978, 61.497, -82.702]
  MoveL 1277 to (0, -7.8, 56.6) mm, rotated rx 180 ry 0 rz 180 deg; joints [-13.166, -51.394, 112.015, 164.973, 61.465, -82.693]
  MoveL 1278 to (-200, -7.8, 56.6) mm, rotated rx 180 ry 0 rz 180 deg; joints [-15.315, -59.455, 128.142, 163.619, 69.479, -84.117]
  MoveL 1279 to (-200, -8.4, 56.6) mm, rotated rx 180 ry 0 rz 180 deg; joints [-15.315, -59.494, 128.141, 163.615, 69.44, -84.104]
  MoveL 1280 to (0, -8.4, 56.6) mm, rotated rx 180 ry 0 rz 180 deg; joints [-13.166, -51.426, 112.014, 164.969, 61.434, -82.683]
  MoveL 1281 to (0, -9, 56.6) mm, rotated rx 180 ry 0 rz 180 deg; joints [-13.166, -51.458, 112.013, 164.964, 61.402, -82.673]
  MoveL 1282 to (-200, -9, 56.6) mm, rotated rx 180 ry 0 rz 180 deg; joints [-15.315, -59.533, 128.139, 163.611, 69.401, -84.092]
  MoveL 1283 to (-200, -9.6, 56.6) mm, rotated rx 180 ry 0 rz 180 deg; joints [-15.315, -59.572, 128.138, 163.606, 69.362, -84.08]
  MoveL 1284 to (0, -9.6, 56.6) mm, rotated rx 180 ry 0 rz 180 deg; joints [-13.166, -51.49, 112.012, 164.959, 61.37, -82.663]
  MoveL 1285 to (0, -10.2, 56.6) mm, rotated rx 180 ry 0 rz 180 deg; joints [-13.166, -51.522, 112.011, 164.955, 61.338, -82.654]
  MoveL 1286 to (-200, -10.2, 56.6) mm, rotated rx 180 ry 0 rz 180 deg; joints [-15.315, -59.611, 128.137, 163.602, 69.324, -84.068]
  MoveL 1287 to (-200, -10.8, 56.6) mm, rotated rx 180 ry 0 rz 180 deg; joints [-15.315, -59.65, 128.136, 163.598, 69.285, -84.056]
  MoveL 1288 to (0, -10.8, 56.6) mm, rotated rx 180 ry 0 rz 180 deg; joints [-13.166, -51.554, 112.01, 164.95, 61.306, -82.644]
  MoveL 1289 to (0, -11.4, 56.6) mm, rotated rx 180 ry 0 rz 180 deg; joints [-13.166, -51.585, 112.008, 164.945, 61.274, -82.634]
